    ELSIF ((x0 = TRUE) AND  (x1 = TRUE) AND  (x2 = FALSE) AND  (t0.Q = FALSE)) THEN 
        cstate58 := 2630; y0 := FALSE; y1 := FALSE; t0_start := FALSE; 
    ELSIF ((x0 = TRUE) AND  (x1 = TRUE) AND  (x2 = FALSE) AND  (t0.Q = TRUE)) THEN 
        cstate58 := 2626; y0 := FALSE; y1 := FALSE; t0_start := FALSE; 
    ELSIF ((x0 = TRUE) AND  (x1 = TRUE) AND  (x2 = TRUE) AND  (t0.Q = FALSE)) THEN 
        cstate58 := 2566; y0 := FALSE; y1 := FALSE; t0_start := TRUE; t0_up := FALSE; 
    ELSIF ((x0 = TRUE) AND  (x1 = TRUE) AND  (x2 = TRUE) AND  (t0.Q = TRUE)) THEN 
        cstate58 := 2562; y0 := FALSE; y1 := FALSE; t0_start := TRUE; t0_up := FALSE; 
    END_IF;
7428:
    IF ((x0 = FALSE) AND  (x1 = FALSE) AND  (x2 = FALSE) AND  (t0.Q = FALSE)) THEN 
        cstate58 := 7428; y0 := FALSE; y1 := FALSE; t0_start := FALSE; 
    ELSIF ((x0 = FALSE) AND  (x1 = FALSE) AND  (x2 = FALSE) AND  (t0.Q = TRUE)) THEN 
        cstate58 := 7370; y0 := FALSE; y1 := TRUE; t0_start := FALSE; 
    ELSIF ((x0 = FALSE) AND  (x1 = FALSE) AND  (x2 = TRUE) AND  (t0.Q = FALSE)) THEN 
        cstate58 := 7492; y0 := FALSE; y1 := FALSE; t0_start := TRUE; t0_up := FALSE; 
    ELSIF ((x0 = FALSE) AND  (x1 = FALSE) AND  (x2 = TRUE) AND  (t0.Q = TRUE)) THEN 
        cstate58 := 7500; y0 := FALSE; y1 := TRUE; t0_start := TRUE; t0_up := FALSE; 
    ELSIF ((x0 = FALSE) AND  (x1 = TRUE) AND  (x2 = FALSE) AND  (t0.Q = FALSE)) THEN 
        cstate58 := 6404; y0 := FALSE; y1 := FALSE; t0_start := FALSE; 
    ELSIF ((x0 = FALSE) AND  (x1 = TRUE) AND  (x2 = FALSE) AND  (t0.Q = TRUE)) THEN 
        cstate58 := 6338; y0 := FALSE; y1 := FALSE; t0_start := FALSE; 
    ELSIF ((x0 = FALSE) AND  (x1 = TRUE) AND  (x2 = TRUE) AND  (t0.Q = FALSE)) THEN 
        cstate58 := 6468; y0 := FALSE; y1 := FALSE; t0_start := TRUE; t0_up := FALSE; 
    ELSIF ((x0 = FALSE) AND  (x1 = TRUE) AND  (x2 = TRUE) AND  (t0.Q = TRUE)) THEN 
        cstate58 := 6466; y0 := FALSE; y1 := FALSE; t0_start := TRUE; t0_up := FALSE; 
    ELSIF ((x0 = TRUE) AND  (x1 = FALSE) AND  (x2 = FALSE) AND  (t0.Q = FALSE)) THEN 
        cstate58 := 5256; y0 := TRUE; y1 := FALSE; t0_start := FALSE; 
    ELSIF ((x0 = TRUE) AND  (x1 = FALSE) AND  (x2 = FALSE) AND  (t0.Q = TRUE)) THEN 
        cstate58 := 5186; y0 := TRUE; y1 := FALSE; t0_start := FALSE; 
    ELSIF ((x0 = TRUE) AND  (x1 = FALSE) AND  (x2 = TRUE) AND  (t0.Q = FALSE)) THEN 
        cstate58 := 3784; y0 := FALSE; y1 := FALSE; t0_start := TRUE; t0_up := FALSE; 
    ELSIF ((x0 = TRUE) AND  (x1 = FALSE) AND  (x2 = TRUE) AND  (t0.Q = TRUE)) THEN 
        cstate58 := 3778; y0 := FALSE; y1 := FALSE; t0_start := TRUE; t0_up := FALSE; 
    ELSIF ((x0 = TRUE) AND  (x1 = TRUE) AND  (x2 = FALSE) AND  (t0.Q = FALSE)) THEN 
        cstate58 := 4742; y0 := TRUE; y1 := FALSE; t0_start := FALSE; 
    ELSIF ((x0 = TRUE) AND  (x1 = TRUE) AND  (x2 = FALSE) AND  (t0.Q = TRUE)) THEN 
        cstate58 := 4674; y0 := TRUE; y1 := FALSE; t0_start := FALSE; 
    ELSIF ((x0 = TRUE) AND  (x1 = TRUE) AND  (x2 = TRUE) AND  (t0.Q = FALSE)) THEN 
        cstate58 := 2566; y0 := FALSE; y1 := FALSE; t0_start := TRUE; t0_up := FALSE; 
    ELSIF ((x0 = TRUE) AND  (x1 = TRUE) AND  (x2 = TRUE) AND  (t0.Q = TRUE)) THEN 
        cstate58 := 2562; y0 := FALSE; y1 := FALSE; t0_start := TRUE; t0_up := FALSE; 
    END_IF;
1304:
    IF ((x0 = FALSE) AND  (x1 = FALSE) AND  (x2 = FALSE) AND  (t0.Q = FALSE)) THEN 
        cstate58 := 1304; y0 := FALSE; y1 := TRUE; t0_start := FALSE; 
    ELSIF ((x0 = FALSE) AND  (x1 = FALSE) AND  (x2 = FALSE) AND  (t0.Q = TRUE)) THEN 
        cstate58 := 1226; y0 := FALSE; y1 := TRUE; t0_start := FALSE; 
    ELSIF ((x0 = FALSE) AND  (x1 = FALSE) AND  (x2 = TRUE) AND  (t0.Q = FALSE)) THEN 
        cstate58 := 1368; y0 := FALSE; y1 := TRUE; t0_start := TRUE; t0_up := FALSE; 
    ELSIF ((x0 = FALSE) AND  (x1 = FALSE) AND  (x2 = TRUE) AND  (t0.Q = TRUE)) THEN 
        cstate58 := 1356; y0 := FALSE; y1 := TRUE; t0_start := TRUE; t0_up := FALSE; 
    ELSIF ((x0 = FALSE) AND  (x1 = TRUE) AND  (x2 = FALSE) AND  (t0.Q = FALSE)) THEN 
        cstate58 := 1284; y0 := FALSE; y1 := FALSE; t0_start := FALSE; 
    ELSIF ((x0 = FALSE) AND  (x1 = TRUE) AND  (x2 = FALSE) AND  (t0.Q = TRUE)) THEN 
        cstate58 := 1218; y0 := FALSE; y1 := FALSE; t0_start := FALSE; 
    ELSIF ((x0 = FALSE) AND  (x1 = TRUE) AND  (x2 = TRUE) AND  (t0.Q = FALSE)) THEN 
        cstate58 := 1348; y0 := FALSE; y1 := FALSE; t0_start := TRUE; t0_up := FALSE; 
    ELSIF ((x0 = FALSE) AND  (x1 = TRUE) AND  (x2 = TRUE) AND  (t0.Q = TRUE)) THEN 
        cstate58 := 1346; y0 := FALSE; y1 := FALSE; t0_start := TRUE; t0_up := FALSE; 
    ELSIF ((x0 = TRUE) AND  (x1 = FALSE) AND  (x2 = FALSE) AND  (t0.Q = FALSE)) THEN 
        cstate58 := 5256; y0 := TRUE; y1 := FALSE; t0_start := FALSE; 
    ELSIF ((x0 = TRUE) AND  (x1 = FALSE) AND  (x2 = FALSE) AND  (t0.Q = TRUE)) THEN 
        cstate58 := 5186; y0 := TRUE; y1 := FALSE; t0_start := FALSE; 
    ELSIF ((x0 = TRUE) AND  (x1 = FALSE) AND  (x2 = TRUE) AND  (t0.Q = FALSE)) THEN 
        cstate58 := 3784; y0 := FALSE; y1 := FALSE; t0_start := TRUE; t0_up := FALSE; 
    ELSIF ((x0 = TRUE) AND  (x1 = FALSE) AND  (x2 = TRUE) AND  (t0.Q = TRUE)) THEN 
        cstate58 := 3778; y0 := FALSE; y1 := FALSE; t0_start := TRUE; t0_up := FALSE; 
    ELSIF ((x0 = TRUE) AND  (x1 = TRUE) AND  (x2 = FALSE) AND  (t0.Q = FALSE)) THEN 
        cstate58 := 4742; y0 := TRUE; y1 := FALSE; t0_start := FALSE; 
    ELSIF ((x0 = TRUE) AND  (x1 = TRUE) AND  (x2 = FALSE) AND  (t0.Q = TRUE)) THEN 
        cstate58 := 4674; y0 := TRUE; y1 := FALSE; t0_start := FALSE; 
    ELSIF ((x0 = TRUE) AND  (x1 = TRUE) AND  (x2 = TRUE) AND  (t0.Q = FALSE)) THEN 
        cstate58 := 2566; y0 := FALSE; y1 := FALSE; t0_start := TRUE; t0_up := FALSE; 
    ELSIF ((x0 = TRUE) AND  (x1 = TRUE) AND  (x2 = TRUE) AND  (t0.Q = TRUE)) THEN 
        cstate58 := 2562; y0 := FALSE; y1 := FALSE; t0_start := TRUE; t0_up := FALSE; 
    END_IF;
2824:
    IF ((x0 = FALSE) AND  (x1 = FALSE) AND  (x2 = FALSE) AND  (t0.Q = FALSE)) THEN 
        cstate58 := 6340; y0 := FALSE; y1 := FALSE; t0_start := FALSE; 
    ELSIF ((x0 = FALSE) AND  (x1 = FALSE) AND  (x2 = FALSE) AND  (t0.Q = TRUE)) THEN 
        cstate58 := 6354; y0 := FALSE; y1 := TRUE; t0_start := FALSE; 
    ELSIF ((x0 = FALSE) AND  (x1 = FALSE) AND  (x2 = TRUE) AND  (t0.Q = FALSE)) THEN 
        cstate58 := 6532; y0 := FALSE; y1 := FALSE; t0_start := FALSE; 
    ELSIF ((x0 = FALSE) AND  (x1 = FALSE) AND  (x2 = TRUE) AND  (t0.Q = TRUE)) THEN 
        cstate58 := 6546; y0 := FALSE; y1 := TRUE; t0_start := FALSE; 
    ELSIF ((x0 = FALSE) AND  (x1 = TRUE) AND  (x2 = FALSE) AND  (t0.Q = FALSE)) THEN 
        cstate58 := 6340; y0 := FALSE; y1 := FALSE; t0_start := FALSE; 
    ELSIF ((x0 = FALSE) AND  (x1 = TRUE) AND  (x2 = FALSE) AND  (t0.Q = TRUE)) THEN 
        cstate58 := 6338; y0 := FALSE; y1 := FALSE; t0_start := FALSE; 
    ELSIF ((x0 = FALSE) AND  (x1 = TRUE) AND  (x2 = TRUE) AND  (t0.Q = FALSE)) THEN 
        cstate58 := 6532; y0 := FALSE; y1 := FALSE; t0_start := FALSE; 
    ELSIF ((x0 = FALSE) AND  (x1 = TRUE) AND  (x2 = TRUE) AND  (t0.Q = TRUE)) THEN 
        cstate58 := 6530; y0 := FALSE; y1 := FALSE; t0_start := FALSE; 
    ELSIF ((x0 = TRUE) AND  (x1 = FALSE) AND  (x2 = FALSE) AND  (t0.Q = FALSE)) THEN 
        cstate58 := 2120; y0 := FALSE; y1 := FALSE; t0_start := FALSE; 
    ELSIF ((x0 = TRUE) AND  (x1 = FALSE) AND  (x2 = FALSE) AND  (t0.Q = TRUE)) THEN 
        cstate58 := 2114; y0 := FALSE; y1 := FALSE; t0_start := FALSE; 
    ELSIF ((x0 = TRUE) AND  (x1 = FALSE) AND  (x2 = TRUE) AND  (t0.Q = FALSE)) THEN 
        cstate58 := 2824; y0 := FALSE; y1 := FALSE; t0_start := FALSE; 
    ELSIF ((x0 = TRUE) AND  (x1 = FALSE) AND  (x2 = TRUE) AND  (t0.Q = TRUE)) THEN 
        cstate58 := 2818; y0 := FALSE; y1 := FALSE; t0_start := FALSE; 
    ELSIF ((x0 = TRUE) AND  (x1 = TRUE) AND  (x2 = FALSE) AND  (t0.Q = FALSE)) THEN 
        cstate58 := 2630; y0 := FALSE; y1 := FALSE; t0_start := FALSE; 
    ELSIF ((x0 = TRUE) AND  (x1 = TRUE) AND  (x2 = FALSE) AND  (t0.Q = TRUE)) THEN 
        cstate58 := 2626; y0 := FALSE; y1 := FALSE; t0_start := FALSE; 
    ELSIF ((x0 = TRUE) AND  (x1 = TRUE) AND  (x2 = TRUE) AND  (t0.Q = FALSE)) THEN 
        cstate58 := 2502; y0 := FALSE; y1 := FALSE; t0_start := FALSE; 
    ELSIF ((x0 = TRUE) AND  (x1 = TRUE) AND  (x2 = TRUE) AND  (t0.Q = TRUE)) THEN 
        cstate58 := 2498; y0 := FALSE; y1 := FALSE; t0_start := FALSE; 
    END_IF;
6480:
    IF ((x0 = FALSE) AND  (x1 = FALSE) AND  (x2 = FALSE) AND  (t0.Q = FALSE)) THEN 
        cstate58 := 6428; y0 := FALSE; y1 := TRUE; t0_start := FALSE; 
    ELSIF ((x0 = FALSE) AND  (x1 = FALSE) AND  (x2 = FALSE) AND  (t0.Q = TRUE)) THEN 
        cstate58 := 6350; y0 := FALSE; y1 := TRUE; t0_start := FALSE; 
    ELSIF ((x0 = FALSE) AND  (x1 = FALSE) AND  (x2 = TRUE) AND  (t0.Q = FALSE)) THEN 
        cstate58 := 6492; y0 := FALSE; y1 := TRUE; t0_start := FALSE; 
    ELSIF ((x0 = FALSE) AND  (x1 = FALSE) AND  (x2 = TRUE) AND  (t0.Q = TRUE)) THEN 
        cstate58 := 6542; y0 := FALSE; y1 := TRUE; t0_start := FALSE; 
    ELSIF ((x0 = FALSE) AND  (x1 = TRUE) AND  (x2 = FALSE) AND  (t0.Q = FALSE)) THEN 
        cstate58 := 6404; y0 := FALSE; y1 := FALSE; t0_start := FALSE; 
    ELSIF ((x0 = FALSE) AND  (x1 = TRUE) AND  (x2 = FALSE) AND  (t0.Q = TRUE)) THEN 
        cstate58 := 6338; y0 := FALSE; y1 := FALSE; t0_start := FALSE; 
    ELSIF ((x0 = FALSE) AND  (x1 = TRUE) AND  (x2 = TRUE) AND  (t0.Q = FALSE)) THEN 
        cstate58 := 6468; y0 := FALSE; y1 := FALSE; t0_start := FALSE; 
    ELSIF ((x0 = FALSE) AND  (x1 = TRUE) AND  (x2 = TRUE) AND  (t0.Q = TRUE)) THEN 
        cstate58 := 6530; y0 := FALSE; y1 := FALSE; t0_start := FALSE; 
    ELSIF ((x0 = TRUE) AND  (x1 = FALSE) AND  (x2 = FALSE) AND  (t0.Q = FALSE)) THEN 
        cstate58 := 4232; y0 := TRUE; y1 := FALSE; t0_start := FALSE; 
    ELSIF ((x0 = TRUE) AND  (x1 = FALSE) AND  (x2 = FALSE) AND  (t0.Q = TRUE)) THEN 
        cstate58 := 4162; y0 := TRUE; y1 := FALSE; t0_start := FALSE; 
    ELSIF ((x0 = TRUE) AND  (x1 = FALSE) AND  (x2 = TRUE) AND  (t0.Q = FALSE)) THEN 
        cstate58 := 2760; y0 := FALSE; y1 := FALSE; t0_start := FALSE; 
    ELSIF ((x0 = TRUE) AND  (x1 = FALSE) AND  (x2 = TRUE) AND  (t0.Q = TRUE)) THEN 
        cstate58 := 2818; y0 := FALSE; y1 := FALSE; t0_start := FALSE; 
    ELSIF ((x0 = TRUE) AND  (x1 = TRUE) AND  (x2 = FALSE) AND  (t0.Q = FALSE)) THEN 
        cstate58 := 4742; y0 := TRUE; y1 := FALSE; t0_start := FALSE; 
    ELSIF ((x0 = TRUE) AND  (x1 = TRUE) AND  (x2 = FALSE) AND  (t0.Q = TRUE)) THEN 
        cstate58 := 4674; y0 := TRUE; y1 := FALSE; t0_start := FALSE; 
    ELSIF ((x0 = TRUE) AND  (x1 = TRUE) AND  (x2 = TRUE) AND  (t0.Q = FALSE)) THEN 
        cstate58 := 2566; y0 := FALSE; y1 := FALSE; t0_start := FALSE; 
    ELSIF ((x0 = TRUE) AND  (x1 = TRUE) AND  (x2 = TRUE) AND  (t0.Q = TRUE)) THEN 
        cstate58 := 2498; y0 := FALSE; y1 := FALSE; t0_start := FALSE; 
    END_IF;
6484:
    IF ((x0 = FALSE) AND  (x1 = FALSE) AND  (x2 = FALSE) AND  (t0.Q = FALSE)) THEN 
        cstate58 := 6432; y0 := FALSE; y1 := TRUE; t0_start := FALSE; 
    ELSIF ((x0 = FALSE) AND  (x1 = FALSE) AND  (x2 = FALSE) AND  (t0.Q = TRUE)) THEN 
        cstate58 := 6354; y0 := FALSE; y1 := TRUE; t0_start := FALSE; 
    ELSIF ((x0 = FALSE) AND  (x1 = FALSE) AND  (x2 = TRUE) AND  (t0.Q = FALSE)) THEN 
        cstate58 := 6496; y0 := FALSE; y1 := TRUE; t0_start := FALSE; 
    ELSIF ((x0 = FALSE) AND  (x1 = FALSE) AND  (x2 = TRUE) AND  (t0.Q = TRUE)) THEN 
        cstate58 := 6546; y0 := FALSE; y1 := TRUE; t0_start := FALSE; 
    ELSIF ((x0 = FALSE) AND  (x1 = TRUE) AND  (x2 = FALSE) AND  (t0.Q = FALSE)) THEN 
        cstate58 := 6404; y0 := FALSE; y1 := FALSE; t0_start := FALSE; 
    ELSIF ((x0 = FALSE) AND  (x1 = TRUE) AND  (x2 = FALSE) AND  (t0.Q = TRUE)) THEN 
        cstate58 := 6338; y0 := FALSE; y1 := FALSE; t0_start := FALSE; 
    ELSIF ((x0 = FALSE) AND  (x1 = TRUE) AND  (x2 = TRUE) AND  (t0.Q = FALSE)) THEN 
        cstate58 := 6468; y0 := FALSE; y1 := FALSE; t0_start := FALSE; 
    ELSIF ((x0 = FALSE) AND  (x1 = TRUE) AND  (x2 = TRUE) AND  (t0.Q = TRUE)) THEN 
        cstate58 := 6530; y0 := FALSE; y1 := FALSE; t0_start := FALSE; 
    ELSIF ((x0 = TRUE) AND  (x1 = FALSE) AND  (x2 = FALSE) AND  (t0.Q = FALSE)) THEN 
        cstate58 := 4232; y0 := TRUE; y1 := FALSE; t0_start := FALSE; 
    ELSIF ((x0 = TRUE) AND  (x1 = FALSE) AND  (x2 = FALSE) AND  (t0.Q = TRUE)) THEN 
        cstate58 := 4162; y0 := TRUE; y1 := FALSE; t0_start := FALSE; 
    ELSIF ((x0 = TRUE) AND  (x1 = FALSE) AND  (x2 = TRUE) AND  (t0.Q = FALSE)) THEN 
        cstate58 := 2760; y0 := FALSE; y1 := FALSE; t0_start := FALSE; 
    ELSIF ((x0 = TRUE) AND  (x1 = FALSE) AND  (x2 = TRUE) AND  (t0.Q = TRUE)) THEN 
        cstate58 := 2818; y0 := FALSE; y1 := FALSE; t0_start := FALSE; 
    ELSIF ((x0 = TRUE) AND  (x1 = TRUE) AND  (x2 = FALSE) AND  (t0.Q = FALSE)) THEN 
        cstate58 := 4742; y0 := TRUE; y1 := FALSE; t0_start := FALSE; 
    ELSIF ((x0 = TRUE) AND  (x1 = TRUE) AND  (x2 = FALSE) AND  (t0.Q = TRUE)) THEN 
        cstate58 := 4674; y0 := TRUE; y1 := FALSE; t0_start := FALSE; 
    ELSIF ((x0 = TRUE) AND  (x1 = TRUE) AND  (x2 = TRUE) AND  (t0.Q = FALSE)) THEN 
        cstate58 := 2566; y0 := FALSE; y1 := FALSE; t0_start := FALSE; 
    ELSIF ((x0 = TRUE) AND  (x1 = TRUE) AND  (x2 = TRUE) AND  (t0.Q = TRUE)) THEN 
        cstate58 := 2498; y0 := FALSE; y1 := FALSE; t0_start := FALSE; 
    END_IF;
2184:
    IF ((x0 = FALSE) AND  (x1 = FALSE) AND  (x2 = FALSE) AND  (t0.Q = FALSE)) THEN 
        cstate58 := 6404; y0 := FALSE; y1 := FALSE; t0_start := FALSE; 
    ELSIF ((x0 = FALSE) AND  (x1 = FALSE) AND  (x2 = FALSE) AND  (t0.Q = TRUE)) THEN 
        cstate58 := 6354; y0 := FALSE; y1 := TRUE; t0_start := FALSE; 
    ELSIF ((x0 = FALSE) AND  (x1 = FALSE) AND  (x2 = TRUE) AND  (t0.Q = FALSE)) THEN 
        cstate58 := 6468; y0 := FALSE; y1 := FALSE; t0_start := TRUE; t0_up := FALSE; 
    ELSIF ((x0 = FALSE) AND  (x1 = FALSE) AND  (x2 = TRUE) AND  (t0.Q = TRUE)) THEN 
        cstate58 := 6484; y0 := FALSE; y1 := TRUE; t0_start := TRUE; t0_up := FALSE; 
    ELSIF ((x0 = FALSE) AND  (x1 = TRUE) AND  (x2 = FALSE) AND  (t0.Q = FALSE)) THEN 
        cstate58 := 6404; y0 := FALSE; y1 := FALSE; t0_start := FALSE; 
    ELSIF ((x0 = FALSE) AND  (x1 = TRUE) AND  (x2 = FALSE) AND  (t0.Q = TRUE)) THEN 
        cstate58 := 6338; y0 := FALSE; y1 := FALSE; t0_start := FALSE; 
    ELSIF ((x0 = FALSE) AND  (x1 = TRUE) AND  (x2 = TRUE) AND  (t0.Q = FALSE)) THEN 
        cstate58 := 6468; y0 := FALSE; y1 := FALSE; t0_start := TRUE; t0_up := FALSE; 
    ELSIF ((x0 = FALSE) AND  (x1 = TRUE) AND  (x2 = TRUE) AND  (t0.Q = TRUE)) THEN 
        cstate58 := 6466; y0 := FALSE; y1 := FALSE; t0_start := TRUE; t0_up := FALSE; 
    ELSIF ((x0 = TRUE) AND  (x1 = FALSE) AND  (x2 = FALSE) AND  (t0.Q = FALSE)) THEN 
        cstate58 := 2184; y0 := FALSE; y1 := FALSE; t0_start := FALSE; 
    ELSIF ((x0 = TRUE) AND  (x1 = FALSE) AND  (x2 = FALSE) AND  (t0.Q = TRUE)) THEN 
        cstate58 := 2114; y0 := FALSE; y1 := FALSE; t0_start := FALSE; 
    ELSIF ((x0 = TRUE) AND  (x1 = FALSE) AND  (x2 = TRUE) AND  (t0.Q = FALSE)) THEN 
        cstate58 := 2760; y0 := FALSE; y1 := FALSE; t0_start := TRUE; t0_up := FALSE; 
    ELSIF ((x0 = TRUE) AND  (x1 = FALSE) AND  (x2 = TRUE) AND  (t0.Q = TRUE)) THEN 
        cstate58 := 2754; y0 := FALSE; y1 := FALSE; t0_start := TRUE; t0_up := FALSE; 
    ELSIF ((x0 = TRUE) AND  (x1 = TRUE) AND  (x2 = FALSE) AND  (t0.Q = FALSE)) THEN 
        cstate58 := 2694; y0 := FALSE; y1 := FALSE; t0_start := FALSE; 
    ELSIF ((x0 = TRUE) AND  (x1 = TRUE) AND  (x2 = FALSE) AND  (t0.Q = TRUE)) THEN 
        cstate58 := 2626; y0 := FALSE; y1 := FALSE; t0_start := FALSE; 
    ELSIF ((x0 = TRUE) AND  (x1 = TRUE) AND  (x2 = TRUE) AND  (t0.Q = FALSE)) THEN 
        cstate58 := 2566; y0 := FALSE; y1 := FALSE; t0_start := TRUE; t0_up := FALSE; 
    ELSIF ((x0 = TRUE) AND  (x1 = TRUE) AND  (x2 = TRUE) AND  (t0.Q = TRUE)) THEN 
        cstate58 := 2562; y0 := FALSE; y1 := FALSE; t0_start := TRUE; t0_up := FALSE; 
    END_IF;
6488:
    IF ((x0 = FALSE) AND  (x1 = FALSE) AND  (x2 = FALSE) AND  (t0.Q = FALSE)) THEN 
        cstate58 := 6424; y0 := FALSE; y1 := TRUE; t0_start := FALSE; 
    ELSIF ((x0 = FALSE) AND  (x1 = FALSE) AND  (x2 = FALSE) AND  (t0.Q = TRUE)) THEN 
        cstate58 := 6346; y0 := FALSE; y1 := TRUE; t0_start := FALSE; 
    ELSIF ((x0 = FALSE) AND  (x1 = FALSE) AND  (x2 = TRUE) AND  (t0.Q = FALSE)) THEN 
        cstate58 := 6488; y0 := FALSE; y1 := TRUE; t0_start := FALSE; 
    ELSIF ((x0 = FALSE) AND  (x1 = FALSE) AND  (x2 = TRUE) AND  (t0.Q = TRUE)) THEN 
        cstate58 := 6538; y0 := FALSE; y1 := TRUE; t0_start := FALSE; 
    ELSIF ((x0 = FALSE) AND  (x1 = TRUE) AND  (x2 = FALSE) AND  (t0.Q = FALSE)) THEN 
        cstate58 := 6404; y0 := FALSE; y1 := FALSE; t0_start := FALSE; 
    ELSIF ((x0 = FALSE) AND  (x1 = TRUE) AND  (x2 = FALSE) AND  (t0.Q = TRUE)) THEN 
        cstate58 := 6338; y0 := FALSE; y1 := FALSE; t0_start := FALSE; 
    ELSIF ((x0 = FALSE) AND  (x1 = TRUE) AND  (x2 = TRUE) AND  (t0.Q = FALSE)) THEN 
        cstate58 := 6468; y0 := FALSE; y1 := FALSE; t0_start := FALSE; 
    ELSIF ((x0 = FALSE) AND  (x1 = TRUE) AND  (x2 = TRUE) AND  (t0.Q = TRUE)) THEN 
        cstate58 := 6530; y0 := FALSE; y1 := FALSE; t0_start := FALSE; 
    ELSIF ((x0 = TRUE) AND  (x1 = FALSE) AND  (x2 = FALSE) AND  (t0.Q = FALSE)) THEN 
        cstate58 := 4232; y0 := TRUE; y1 := FALSE; t0_start := FALSE; 
    ELSIF ((x0 = TRUE) AND  (x1 = FALSE) AND  (x2 = FALSE) AND  (t0.Q = TRUE)) THEN 
        cstate58 := 4162; y0 := TRUE; y1 := FALSE; t0_start := FALSE; 
    ELSIF ((x0 = TRUE) AND  (x1 = FALSE) AND  (x2 = TRUE) AND  (t0.Q = FALSE)) THEN 
        cstate58 := 2760; y0 := FALSE; y1 := FALSE; t0_start := FALSE; 
    ELSIF ((x0 = TRUE) AND  (x1 = FALSE) AND  (x2 = TRUE) AND  (t0.Q = TRUE)) THEN 
        cstate58 := 2818; y0 := FALSE; y1 := FALSE; t0_start := FALSE; 
    ELSIF ((x0 = TRUE) AND  (x1 = TRUE) AND  (x2 = FALSE) AND  (t0.Q = FALSE)) THEN 
        cstate58 := 4742; y0 := TRUE; y1 := FALSE; t0_start := FALSE; 
    ELSIF ((x0 = TRUE) AND  (x1 = TRUE) AND  (x2 = FALSE) AND  (t0.Q = TRUE)) THEN 
        cstate58 := 4674; y0 := TRUE; y1 := FALSE; t0_start := FALSE; 
    ELSIF ((x0 = TRUE) AND  (x1 = TRUE) AND  (x2 = TRUE) AND  (t0.Q = FALSE)) THEN 
        cstate58 := 2566; y0 := FALSE; y1 := FALSE; t0_start := FALSE; 
    ELSIF ((x0 = TRUE) AND  (x1 = TRUE) AND  (x2 = TRUE) AND  (t0.Q = TRUE)) THEN 
        cstate58 := 2498; y0 := FALSE; y1 := FALSE; t0_start := FALSE; 
    END_IF;
6466:
    IF ((x0 = FALSE) AND  (x1 = FALSE) AND  (x2 = FALSE) AND  (t0.Q = FALSE)) THEN 
        cstate58 := 6404; y0 := FALSE; y1 := FALSE; t0_start := FALSE; 
    ELSIF ((x0 = FALSE) AND  (x1 = FALSE) AND  (x2 = FALSE) AND  (t0.Q = TRUE)) THEN 
        cstate58 := 6338; y0 := FALSE; y1 := FALSE; t0_start := FALSE; 
    ELSIF ((x0 = FALSE) AND  (x1 = FALSE) AND  (x2 = TRUE) AND  (t0.Q = FALSE)) THEN 
        cstate58 := 6468; y0 := FALSE; y1 := FALSE; t0_start := FALSE; 
    ELSIF ((x0 = FALSE) AND  (x1 = FALSE) AND  (x2 = TRUE) AND  (t0.Q = TRUE)) THEN 
        cstate58 := 6530; y0 := FALSE; y1 := FALSE; t0_start := FALSE; 
    ELSIF ((x0 = FALSE) AND  (x1 = TRUE) AND  (x2 = FALSE) AND  (t0.Q = FALSE)) THEN 
        cstate58 := 6404; y0 := FALSE; y1 := FALSE; t0_start := FALSE; 
    ELSIF ((x0 = FALSE) AND  (x1 = TRUE) AND  (x2 = FALSE) AND  (t0.Q = TRUE)) THEN 
        cstate58 := 6338; y0 := FALSE; y1 := FALSE; t0_start := FALSE; 
    ELSIF ((x0 = FALSE) AND  (x1 = TRUE) AND  (x2 = TRUE) AND  (t0.Q = FALSE)) THEN 
        cstate58 := 6468; y0 := FALSE; y1 := FALSE; t0_start := FALSE; 
    ELSIF ((x0 = FALSE) AND  (x1 = TRUE) AND  (x2 = TRUE) AND  (t0.Q = TRUE)) THEN 
        cstate58 := 6530; y0 := FALSE; y1 := FALSE; t0_start := FALSE; 
    ELSIF ((x0 = TRUE) AND  (x1 = FALSE) AND  (x2 = FALSE) AND  (t0.Q = FALSE)) THEN 
        cstate58 := 4232; y0 := TRUE; y1 := FALSE; t0_start := FALSE; 
    ELSIF ((x0 = TRUE) AND  (x1 = FALSE) AND  (x2 = FALSE) AND  (t0.Q = TRUE)) THEN 
        cstate58 := 4162; y0 := TRUE; y1 := FALSE; t0_start := FALSE; 
    ELSIF ((x0 = TRUE) AND  (x1 = FALSE) AND  (x2 = TRUE) AND  (t0.Q = FALSE)) THEN 
        cstate58 := 2760; y0 := FALSE; y1 := FALSE; t0_start := FALSE; 
    ELSIF ((x0 = TRUE) AND  (x1 = FALSE) AND  (x2 = TRUE) AND  (t0.Q = TRUE)) THEN 
        cstate58 := 2818; y0 := FALSE; y1 := FALSE; t0_start := FALSE; 
    ELSIF ((x0 = TRUE) AND  (x1 = TRUE) AND  (x2 = FALSE) AND  (t0.Q = FALSE)) THEN 
        cstate58 := 4742; y0 := TRUE; y1 := FALSE; t0_start := FALSE; 
    ELSIF ((x0 = TRUE) AND  (x1 = TRUE) AND  (x2 = FALSE) AND  (t0.Q = TRUE)) THEN 
        cstate58 := 4674; y0 := TRUE; y1 := FALSE; t0_start := FALSE; 
    ELSIF ((x0 = TRUE) AND  (x1 = TRUE) AND  (x2 = TRUE) AND  (t0.Q = FALSE)) THEN 
        cstate58 := 2566; y0 := FALSE; y1 := FALSE; t0_start := FALSE; 
    ELSIF ((x0 = TRUE) AND  (x1 = TRUE) AND  (x2 = TRUE) AND  (t0.Q = TRUE)) THEN 
        cstate58 := 2498; y0 := FALSE; y1 := FALSE; t0_start := FALSE; 
    END_IF;
9410:
    IF ((x0 = FALSE) AND  (x1 = FALSE) AND  (x2 = FALSE) AND  (t0.Q = FALSE)) THEN 
        cstate58 := 9412; y0 := TRUE; y1 := FALSE; t0_start := FALSE; 
    ELSIF ((x0 = FALSE) AND  (x1 = FALSE) AND  (x2 = FALSE) AND  (t0.Q = TRUE)) THEN 
        cstate58 := 9410; y0 := TRUE; y1 := FALSE; t0_start := FALSE; 
    ELSIF ((x0 = FALSE) AND  (x1 = FALSE) AND  (x2 = TRUE) AND  (t0.Q = FALSE)) THEN 
        cstate58 := 7492; y0 := FALSE; y1 := FALSE; t0_start := TRUE; t0_up := FALSE; 
    ELSIF ((x0 = FALSE) AND  (x1 = FALSE) AND  (x2 = TRUE) AND  (t0.Q = TRUE)) THEN 
        cstate58 := 7490; y0 := FALSE; y1 := FALSE; t0_start := TRUE; t0_up := FALSE; 
    ELSIF ((x0 = FALSE) AND  (x1 = TRUE) AND  (x2 = FALSE) AND  (t0.Q = FALSE)) THEN 
        cstate58 := 8388; y0 := TRUE; y1 := FALSE; t0_start := FALSE; 
    ELSIF ((x0 = FALSE) AND  (x1 = TRUE) AND  (x2 = FALSE) AND  (t0.Q = TRUE)) THEN 
        cstate58 := 8386; y0 := TRUE; y1 := FALSE; t0_start := FALSE; 
    ELSIF ((x0 = FALSE) AND  (x1 = TRUE) AND  (x2 = TRUE) AND  (t0.Q = FALSE)) THEN 
        cstate58 := 6468; y0 := FALSE; y1 := FALSE; t0_start := TRUE; t0_up := FALSE; 
    ELSIF ((x0 = FALSE) AND  (x1 = TRUE) AND  (x2 = TRUE) AND  (t0.Q = TRUE)) THEN 
        cstate58 := 6466; y0 := FALSE; y1 := FALSE; t0_start := TRUE; t0_up := FALSE; 
    ELSIF ((x0 = TRUE) AND  (x1 = FALSE) AND  (x2 = FALSE) AND  (t0.Q = FALSE)) THEN 
        cstate58 := 5192; y0 := TRUE; y1 := FALSE; t0_start := FALSE; 
    ELSIF ((x0 = TRUE) AND  (x1 = FALSE) AND  (x2 = FALSE) AND  (t0.Q = TRUE)) THEN 
        cstate58 := 5186; y0 := TRUE; y1 := FALSE; t0_start := FALSE; 
    ELSIF ((x0 = TRUE) AND  (x1 = FALSE) AND  (x2 = TRUE) AND  (t0.Q = FALSE)) THEN 
        cstate58 := 3784; y0 := FALSE; y1 := FALSE; t0_start := TRUE; t0_up := FALSE; 
    ELSIF ((x0 = TRUE) AND  (x1 = FALSE) AND  (x2 = TRUE) AND  (t0.Q = TRUE)) THEN 
        cstate58 := 3778; y0 := FALSE; y1 := FALSE; t0_start := TRUE; t0_up := FALSE; 
    ELSIF ((x0 = TRUE) AND  (x1 = TRUE) AND  (x2 = FALSE) AND  (t0.Q = FALSE)) THEN 
        cstate58 := 4678; y0 := TRUE; y1 := FALSE; t0_start := FALSE; 
    ELSIF ((x0 = TRUE) AND  (x1 = TRUE) AND  (x2 = FALSE) AND  (t0.Q = TRUE)) THEN 
        cstate58 := 4674; y0 := TRUE; y1 := FALSE; t0_start := FALSE; 
    ELSIF ((x0 = TRUE) AND  (x1 = TRUE) AND  (x2 = TRUE) AND  (t0.Q = FALSE)) THEN 
        cstate58 := 2566; y0 := FALSE; y1 := FALSE; t0_start := TRUE; t0_up := FALSE; 
    ELSIF ((x0 = TRUE) AND  (x1 = TRUE) AND  (x2 = TRUE) AND  (t0.Q = TRUE)) THEN 
        cstate58 := 2562; y0 := FALSE; y1 := FALSE; t0_start := TRUE; t0_up := FALSE; 
    END_IF;
2818:
    IF ((x0 = FALSE) AND  (x1 = FALSE) AND  (x2 = FALSE) AND  (t0.Q = FALSE)) THEN 
        cstate58 := 6340; y0 := FALSE; y1 := FALSE; t0_start := FALSE; 
    ELSIF ((x0 = FALSE) AND  (x1 = FALSE) AND  (x2 = FALSE) AND  (t0.Q = TRUE)) THEN 
        cstate58 := 6338; y0 := FALSE; y1 := FALSE; t0_start := FALSE; 
    ELSIF ((x0 = FALSE) AND  (x1 = FALSE) AND  (x2 = TRUE) AND  (t0.Q = FALSE)) THEN 
        cstate58 := 6532; y0 := FALSE; y1 := FALSE; t0_start := FALSE; 
    ELSIF ((x0 = FALSE) AND  (x1 = FALSE) AND  (x2 = TRUE) AND  (t0.Q = TRUE)) THEN 
        cstate58 := 6530; y0 := FALSE; y1 := FALSE; t0_start := FALSE; 
    ELSIF ((x0 = FALSE) AND  (x1 = TRUE) AND  (x2 = FALSE) AND  (t0.Q = FALSE)) THEN 
        cstate58 := 6340; y0 := FALSE; y1 := FALSE; t0_start := FALSE; 
    ELSIF ((x0 = FALSE) AND  (x1 = TRUE) AND  (x2 = FALSE) AND  (t0.Q = TRUE)) THEN 
        cstate58 := 6338; y0 := FALSE; y1 := FALSE; t0_start := FALSE; 
    ELSIF ((x0 = FALSE) AND  (x1 = TRUE) AND  (x2 = TRUE) AND  (t0.Q = FALSE)) THEN 
        cstate58 := 6532; y0 := FALSE; y1 := FALSE; t0_start := FALSE; 
    ELSIF ((x0 = FALSE) AND  (x1 = TRUE) AND  (x2 = TRUE) AND  (t0.Q = TRUE)) THEN 
        cstate58 := 6530; y0 := FALSE; y1 := FALSE; t0_start := FALSE; 
    ELSIF ((x0 = TRUE) AND  (x1 = FALSE) AND  (x2 = FALSE) AND  (t0.Q = FALSE)) THEN 
        cstate58 := 2120; y0 := FALSE; y1 := FALSE; t0_start := FALSE; 
    ELSIF ((x0 = TRUE) AND  (x1 = FALSE) AND  (x2 = FALSE) AND  (t0.Q = TRUE)) THEN 
        cstate58 := 2114; y0 := FALSE; y1 := FALSE; t0_start := FALSE; 
    ELSIF ((x0 = TRUE) AND  (x1 = FALSE) AND  (x2 = TRUE) AND  (t0.Q = FALSE)) THEN 
        cstate58 := 2824; y0 := FALSE; y1 := FALSE; t0_start := FALSE; 
    ELSIF ((x0 = TRUE) AND  (x1 = FALSE) AND  (x2 = TRUE) AND  (t0.Q = TRUE)) THEN 
        cstate58 := 2818; y0 := FALSE; y1 := FALSE; t0_start := FALSE; 
    ELSIF ((x0 = TRUE) AND  (x1 = TRUE) AND  (x2 = FALSE) AND  (t0.Q = FALSE)) THEN 
        cstate58 := 2630; y0 := FALSE; y1 := FALSE; t0_start := FALSE; 
    ELSIF ((x0 = TRUE) AND  (x1 = TRUE) AND  (x2 = FALSE) AND  (t0.Q = TRUE)) THEN 
        cstate58 := 2626; y0 := FALSE; y1 := FALSE; t0_start := FALSE; 
    ELSIF ((x0 = TRUE) AND  (x1 = TRUE) AND  (x2 = TRUE) AND  (t0.Q = FALSE)) THEN 
        cstate58 := 2502; y0 := FALSE; y1 := FALSE; t0_start := FALSE; 
    ELSIF ((x0 = TRUE) AND  (x1 = TRUE) AND  (x2 = TRUE) AND  (t0.Q = TRUE)) THEN 
        cstate58 := 2498; y0 := FALSE; y1 := FALSE; t0_start := FALSE; 
    END_IF;
9412:
    IF ((x0 = FALSE) AND  (x1 = FALSE) AND  (x2 = FALSE) AND  (t0.Q = FALSE)) THEN 
        cstate58 := 9412; y0 := TRUE; y1 := FALSE; t0_start := FALSE; 
    ELSIF ((x0 = FALSE) AND  (x1 = FALSE) AND  (x2 = FALSE) AND  (t0.Q = TRUE)) THEN 
        cstate58 := 9410; y0 := TRUE; y1 := FALSE; t0_start := FALSE; 
    ELSIF ((x0 = FALSE) AND  (x1 = FALSE) AND  (x2 = TRUE) AND  (t0.Q = FALSE)) THEN 
        cstate58 := 7492; y0 := FALSE; y1 := FALSE; t0_start := TRUE; t0_up := FALSE; 
    ELSIF ((x0 = FALSE) AND  (x1 = FALSE) AND  (x2 = TRUE) AND  (t0.Q = TRUE)) THEN 
        cstate58 := 7500; y0 := FALSE; y1 := TRUE; t0_start := TRUE; t0_up := FALSE; 
    ELSIF ((x0 = FALSE) AND  (x1 = TRUE) AND  (x2 = FALSE) AND  (t0.Q = FALSE)) THEN 
        cstate58 := 8388; y0 := TRUE; y1 := FALSE; t0_start := FALSE; 
    ELSIF ((x0 = FALSE) AND  (x1 = TRUE) AND  (x2 = FALSE) AND  (t0.Q = TRUE)) THEN 
        cstate58 := 8386; y0 := TRUE; y1 := FALSE; t0_start := FALSE; 
    ELSIF ((x0 = FALSE) AND  (x1 = TRUE) AND  (x2 = TRUE) AND  (t0.Q = FALSE)) THEN 
        cstate58 := 6468; y0 := FALSE; y1 := FALSE; t0_start := TRUE; t0_up := FALSE; 
    ELSIF ((x0 = FALSE) AND  (x1 = TRUE) AND  (x2 = TRUE) AND  (t0.Q = TRUE)) THEN 
        cstate58 := 6466; y0 := FALSE; y1 := FALSE; t0_start := TRUE; t0_up := FALSE; 
    ELSIF ((x0 = TRUE) AND  (x1 = FALSE) AND  (x2 = FALSE) AND  (t0.Q = FALSE)) THEN 
        cstate58 := 5192; y0 := TRUE; y1 := FALSE; t0_start := FALSE; 
    ELSIF ((x0 = TRUE) AND  (x1 = FALSE) AND  (x2 = FALSE) AND  (t0.Q = TRUE)) THEN 
        cstate58 := 5186; y0 := TRUE; y1 := FALSE; t0_start := FALSE; 
    ELSIF ((x0 = TRUE) AND  (x1 = FALSE) AND  (x2 = TRUE) AND  (t0.Q = FALSE)) THEN 
        cstate58 := 3784; y0 := FALSE; y1 := FALSE; t0_start := TRUE; t0_up := FALSE; 
    ELSIF ((x0 = TRUE) AND  (x1 = FALSE) AND  (x2 = TRUE) AND  (t0.Q = TRUE)) THEN 
        cstate58 := 3778; y0 := FALSE; y1 := FALSE; t0_start := TRUE; t0_up := FALSE; 
    ELSIF ((x0 = TRUE) AND  (x1 = TRUE) AND  (x2 = FALSE) AND  (t0.Q = FALSE)) THEN 
        cstate58 := 4678; y0 := TRUE; y1 := FALSE; t0_start := FALSE; 
    ELSIF ((x0 = TRUE) AND  (x1 = TRUE) AND  (x2 = FALSE) AND  (t0.Q = TRUE)) THEN 
        cstate58 := 4674; y0 := TRUE; y1 := FALSE; t0_start := FALSE; 
    ELSIF ((x0 = TRUE) AND  (x1 = TRUE) AND  (x2 = TRUE) AND  (t0.Q = FALSE)) THEN 
        cstate58 := 2566; y0 := FALSE; y1 := FALSE; t0_start := TRUE; t0_up := FALSE; 
    ELSIF ((x0 = TRUE) AND  (x1 = TRUE) AND  (x2 = TRUE) AND  (t0.Q = TRUE)) THEN 
        cstate58 := 2562; y0 := FALSE; y1 := FALSE; t0_start := TRUE; t0_up := FALSE; 
    END_IF;
7456:
    IF ((x0 = FALSE) AND  (x1 = FALSE) AND  (x2 = FALSE) AND  (t0.Q = FALSE)) THEN 
        cstate58 := 7456; y0 := FALSE; y1 := TRUE; t0_start := FALSE; 
    ELSIF ((x0 = FALSE) AND  (x1 = FALSE) AND  (x2 = FALSE) AND  (t0.Q = TRUE)) THEN 
        cstate58 := 7378; y0 := FALSE; y1 := TRUE; t0_start := FALSE; 
    ELSIF ((x0 = FALSE) AND  (x1 = FALSE) AND  (x2 = TRUE) AND  (t0.Q = FALSE)) THEN 
        cstate58 := 7520; y0 := FALSE; y1 := TRUE; t0_start := TRUE; t0_up := FALSE; 
    ELSIF ((x0 = FALSE) AND  (x1 = FALSE) AND  (x2 = TRUE) AND  (t0.Q = TRUE)) THEN 
        cstate58 := 7508; y0 := FALSE; y1 := TRUE; t0_start := TRUE; t0_up := FALSE; 
    ELSIF ((x0 = FALSE) AND  (x1 = TRUE) AND  (x2 = FALSE) AND  (t0.Q = FALSE)) THEN 
        cstate58 := 6404; y0 := FALSE; y1 := FALSE; t0_start := FALSE; 
    ELSIF ((x0 = FALSE) AND  (x1 = TRUE) AND  (x2 = FALSE) AND  (t0.Q = TRUE)) THEN 
        cstate58 := 6338; y0 := FALSE; y1 := FALSE; t0_start := FALSE; 
    ELSIF ((x0 = FALSE) AND  (x1 = TRUE) AND  (x2 = TRUE) AND  (t0.Q = FALSE)) THEN 
        cstate58 := 6468; y0 := FALSE; y1 := FALSE; t0_start := TRUE; t0_up := FALSE; 
    ELSIF ((x0 = FALSE) AND  (x1 = TRUE) AND  (x2 = TRUE) AND  (t0.Q = TRUE)) THEN 
        cstate58 := 6466; y0 := FALSE; y1 := FALSE; t0_start := TRUE; t0_up := FALSE; 
    ELSIF ((x0 = TRUE) AND  (x1 = FALSE) AND  (x2 = FALSE) AND  (t0.Q = FALSE)) THEN 
        cstate58 := 5256; y0 := TRUE; y1 := FALSE; t0_start := FALSE; 
    ELSIF ((x0 = TRUE) AND  (x1 = FALSE) AND  (x2 = FALSE) AND  (t0.Q = TRUE)) THEN 
        cstate58 := 5186; y0 := TRUE; y1 := FALSE; t0_start := FALSE; 
    ELSIF ((x0 = TRUE) AND  (x1 = FALSE) AND  (x2 = TRUE) AND  (t0.Q = FALSE)) THEN 
        cstate58 := 3784; y0 := FALSE; y1 := FALSE; t0_start := TRUE; t0_up := FALSE; 
    ELSIF ((x0 = TRUE) AND  (x1 = FALSE) AND  (x2 = TRUE) AND  (t0.Q = TRUE)) THEN 
        cstate58 := 3778; y0 := FALSE; y1 := FALSE; t0_start := TRUE; t0_up := FALSE; 
    ELSIF ((x0 = TRUE) AND  (x1 = TRUE) AND  (x2 = FALSE) AND  (t0.Q = FALSE)) THEN 
        cstate58 := 4742; y0 := TRUE; y1 := FALSE; t0_start := FALSE; 
    ELSIF ((x0 = TRUE) AND  (x1 = TRUE) AND  (x2 = FALSE) AND  (t0.Q = TRUE)) THEN 
        cstate58 := 4674; y0 := TRUE; y1 := FALSE; t0_start := FALSE; 
    ELSIF ((x0 = TRUE) AND  (x1 = TRUE) AND  (x2 = TRUE) AND  (t0.Q = FALSE)) THEN 
        cstate58 := 2566; y0 := FALSE; y1 := FALSE; t0_start := TRUE; t0_up := FALSE; 
    ELSIF ((x0 = TRUE) AND  (x1 = TRUE) AND  (x2 = TRUE) AND  (t0.Q = TRUE)) THEN 
        cstate58 := 2562; y0 := FALSE; y1 := FALSE; t0_start := TRUE; t0_up := FALSE; 
    END_IF;
7448:
    IF ((x0 = FALSE) AND  (x1 = FALSE) AND  (x2 = FALSE) AND  (t0.Q = FALSE)) THEN 
        cstate58 := 7448; y0 := FALSE; y1 := TRUE; t0_start := FALSE; 
    ELSIF ((x0 = FALSE) AND  (x1 = FALSE) AND  (x2 = FALSE) AND  (t0.Q = TRUE)) THEN 
        cstate58 := 7370; y0 := FALSE; y1 := TRUE; t0_start := FALSE; 
    ELSIF ((x0 = FALSE) AND  (x1 = FALSE) AND  (x2 = TRUE) AND  (t0.Q = FALSE)) THEN 
        cstate58 := 7512; y0 := FALSE; y1 := TRUE; t0_start := TRUE; t0_up := FALSE; 
    ELSIF ((x0 = FALSE) AND  (x1 = FALSE) AND  (x2 = TRUE) AND  (t0.Q = TRUE)) THEN 
        cstate58 := 7500; y0 := FALSE; y1 := TRUE; t0_start := TRUE; t0_up := FALSE; 
    ELSIF ((x0 = FALSE) AND  (x1 = TRUE) AND  (x2 = FALSE) AND  (t0.Q = FALSE)) THEN 
        cstate58 := 6404; y0 := FALSE; y1 := FALSE; t0_start := FALSE; 
    ELSIF ((x0 = FALSE) AND  (x1 = TRUE) AND  (x2 = FALSE) AND  (t0.Q = TRUE)) THEN 
        cstate58 := 6338; y0 := FALSE; y1 := FALSE; t0_start := FALSE; 
    ELSIF ((x0 = FALSE) AND  (x1 = TRUE) AND  (x2 = TRUE) AND  (t0.Q = FALSE)) THEN 
        cstate58 := 6468; y0 := FALSE; y1 := FALSE; t0_start := TRUE; t0_up := FALSE; 
    ELSIF ((x0 = FALSE) AND  (x1 = TRUE) AND  (x2 = TRUE) AND  (t0.Q = TRUE)) THEN 
        cstate58 := 6466; y0 := FALSE; y1 := FALSE; t0_start := TRUE; t0_up := FALSE; 
    ELSIF ((x0 = TRUE) AND  (x1 = FALSE) AND  (x2 = FALSE) AND  (t0.Q = FALSE)) THEN 
        cstate58 := 5256; y0 := TRUE; y1 := FALSE; t0_start := FALSE; 
    ELSIF ((x0 = TRUE) AND  (x1 = FALSE) AND  (x2 = FALSE) AND  (t0.Q = TRUE)) THEN 
        cstate58 := 5186; y0 := TRUE; y1 := FALSE; t0_start := FALSE; 
    ELSIF ((x0 = TRUE) AND  (x1 = FALSE) AND  (x2 = TRUE) AND  (t0.Q = FALSE)) THEN 
        cstate58 := 3784; y0 := FALSE; y1 := FALSE; t0_start := TRUE; t0_up := FALSE; 
    ELSIF ((x0 = TRUE) AND  (x1 = FALSE) AND  (x2 = TRUE) AND  (t0.Q = TRUE)) THEN 
        cstate58 := 3778; y0 := FALSE; y1 := FALSE; t0_start := TRUE; t0_up := FALSE; 
    ELSIF ((x0 = TRUE) AND  (x1 = TRUE) AND  (x2 = FALSE) AND  (t0.Q = FALSE)) THEN 
        cstate58 := 4742; y0 := TRUE; y1 := FALSE; t0_start := FALSE; 
    ELSIF ((x0 = TRUE) AND  (x1 = TRUE) AND  (x2 = FALSE) AND  (t0.Q = TRUE)) THEN 
        cstate58 := 4674; y0 := TRUE; y1 := FALSE; t0_start := FALSE; 
    ELSIF ((x0 = TRUE) AND  (x1 = TRUE) AND  (x2 = TRUE) AND  (t0.Q = FALSE)) THEN 
        cstate58 := 2566; y0 := FALSE; y1 := FALSE; t0_start := TRUE; t0_up := FALSE; 
    ELSIF ((x0 = TRUE) AND  (x1 = TRUE) AND  (x2 = TRUE) AND  (t0.Q = TRUE)) THEN 
        cstate58 := 2562; y0 := FALSE; y1 := FALSE; t0_start := TRUE; t0_up := FALSE; 
    END_IF;
3778:
    IF ((x0 = FALSE) AND  (x1 = FALSE) AND  (x2 = FALSE) AND  (t0.Q = FALSE)) THEN 
        cstate58 := 7428; y0 := FALSE; y1 := FALSE; t0_start := FALSE; 
    ELSIF ((x0 = FALSE) AND  (x1 = FALSE) AND  (x2 = FALSE) AND  (t0.Q = TRUE)) THEN 
        cstate58 := 7362; y0 := FALSE; y1 := FALSE; t0_start := FALSE; 
    ELSIF ((x0 = FALSE) AND  (x1 = FALSE) AND  (x2 = TRUE) AND  (t0.Q = FALSE)) THEN 
        cstate58 := 7492; y0 := FALSE; y1 := FALSE; t0_start := FALSE; 
    ELSIF ((x0 = FALSE) AND  (x1 = FALSE) AND  (x2 = TRUE) AND  (t0.Q = TRUE)) THEN 
        cstate58 := 7554; y0 := FALSE; y1 := FALSE; t0_start := FALSE; 
    ELSIF ((x0 = FALSE) AND  (x1 = TRUE) AND  (x2 = FALSE) AND  (t0.Q = FALSE)) THEN 
        cstate58 := 6404; y0 := FALSE; y1 := FALSE; t0_start := FALSE; 
    ELSIF ((x0 = FALSE) AND  (x1 = TRUE) AND  (x2 = FALSE) AND  (t0.Q = TRUE)) THEN 
        cstate58 := 6338; y0 := FALSE; y1 := FALSE; t0_start := FALSE; 
    ELSIF ((x0 = FALSE) AND  (x1 = TRUE) AND  (x2 = TRUE) AND  (t0.Q = FALSE)) THEN 
        cstate58 := 6468; y0 := FALSE; y1 := FALSE; t0_start := FALSE; 
    ELSIF ((x0 = FALSE) AND  (x1 = TRUE) AND  (x2 = TRUE) AND  (t0.Q = TRUE)) THEN 
        cstate58 := 6530; y0 := FALSE; y1 := FALSE; t0_start := FALSE; 
    ELSIF ((x0 = TRUE) AND  (x1 = FALSE) AND  (x2 = FALSE) AND  (t0.Q = FALSE)) THEN 
        cstate58 := 3208; y0 := FALSE; y1 := FALSE; t0_start := FALSE; 
    ELSIF ((x0 = TRUE) AND  (x1 = FALSE) AND  (x2 = FALSE) AND  (t0.Q = TRUE)) THEN 
        cstate58 := 3138; y0 := FALSE; y1 := FALSE; t0_start := FALSE; 
    ELSIF ((x0 = TRUE) AND  (x1 = FALSE) AND  (x2 = TRUE) AND  (t0.Q = FALSE)) THEN 
        cstate58 := 3784; y0 := FALSE; y1 := FALSE; t0_start := FALSE; 
    ELSIF ((x0 = TRUE) AND  (x1 = FALSE) AND  (x2 = TRUE) AND  (t0.Q = TRUE)) THEN 
        cstate58 := 3842; y0 := FALSE; y1 := FALSE; t0_start := FALSE; 
    ELSIF ((x0 = TRUE) AND  (x1 = TRUE) AND  (x2 = FALSE) AND  (t0.Q = FALSE)) THEN 
        cstate58 := 2694; y0 := FALSE; y1 := FALSE; t0_start := FALSE; 
    ELSIF ((x0 = TRUE) AND  (x1 = TRUE) AND  (x2 = FALSE) AND  (t0.Q = TRUE)) THEN 
        cstate58 := 2626; y0 := FALSE; y1 := FALSE; t0_start := FALSE; 
    ELSIF ((x0 = TRUE) AND  (x1 = TRUE) AND  (x2 = TRUE) AND  (t0.Q = FALSE)) THEN 
        cstate58 := 2566; y0 := FALSE; y1 := FALSE; t0_start := FALSE; 
    ELSIF ((x0 = TRUE) AND  (x1 = TRUE) AND  (x2 = TRUE) AND  (t0.Q = TRUE)) THEN 
        cstate58 := 2498; y0 := FALSE; y1 := FALSE; t0_start := FALSE; 
    END_IF;
7390:
    IF ((x0 = FALSE) AND  (x1 = FALSE) AND  (x2 = FALSE) AND  (t0.Q = FALSE)) THEN 
        cstate58 := 7390; y0 := FALSE; y1 := TRUE; t0_start := FALSE; 
    ELSIF ((x0 = FALSE) AND  (x1 = FALSE) AND  (x2 = FALSE) AND  (t0.Q = TRUE)) THEN 
        cstate58 := 7378; y0 := FALSE; y1 := TRUE; t0_start := FALSE; 
    ELSIF ((x0 = FALSE) AND  (x1 = FALSE) AND  (x2 = TRUE) AND  (t0.Q = FALSE)) THEN 
        cstate58 := 7520; y0 := FALSE; y1 := TRUE; t0_start := TRUE; t0_up := FALSE; 
    ELSIF ((x0 = FALSE) AND  (x1 = FALSE) AND  (x2 = TRUE) AND  (t0.Q = TRUE)) THEN 
        cstate58 := 7508; y0 := FALSE; y1 := TRUE; t0_start := TRUE; t0_up := FALSE; 
    ELSIF ((x0 = FALSE) AND  (x1 = TRUE) AND  (x2 = FALSE) AND  (t0.Q = FALSE)) THEN 
        cstate58 := 6340; y0 := FALSE; y1 := FALSE; t0_start := FALSE; 
    ELSIF ((x0 = FALSE) AND  (x1 = TRUE) AND  (x2 = FALSE) AND  (t0.Q = TRUE)) THEN 
        cstate58 := 6338; y0 := FALSE; y1 := FALSE; t0_start := FALSE; 
    ELSIF ((x0 = FALSE) AND  (x1 = TRUE) AND  (x2 = TRUE) AND  (t0.Q = FALSE)) THEN 
        cstate58 := 6468; y0 := FALSE; y1 := FALSE; t0_start := TRUE; t0_up := FALSE; 
    ELSIF ((x0 = FALSE) AND  (x1 = TRUE) AND  (x2 = TRUE) AND  (t0.Q = TRUE)) THEN 
        cstate58 := 6466; y0 := FALSE; y1 := FALSE; t0_start := TRUE; t0_up := FALSE; 
    ELSIF ((x0 = TRUE) AND  (x1 = FALSE) AND  (x2 = FALSE) AND  (t0.Q = FALSE)) THEN 
        cstate58 := 5192; y0 := TRUE; y1 := FALSE; t0_start := FALSE; 
    ELSIF ((x0 = TRUE) AND  (x1 = FALSE) AND  (x2 = FALSE) AND  (t0.Q = TRUE)) THEN 
        cstate58 := 5186; y0 := TRUE; y1 := FALSE; t0_start := FALSE; 
    ELSIF ((x0 = TRUE) AND  (x1 = FALSE) AND  (x2 = TRUE) AND  (t0.Q = FALSE)) THEN 
        cstate58 := 3784; y0 := FALSE; y1 := FALSE; t0_start := TRUE; t0_up := FALSE; 
    ELSIF ((x0 = TRUE) AND  (x1 = FALSE) AND  (x2 = TRUE) AND  (t0.Q = TRUE)) THEN 
        cstate58 := 3778; y0 := FALSE; y1 := FALSE; t0_start := TRUE; t0_up := FALSE; 
    ELSIF ((x0 = TRUE) AND  (x1 = TRUE) AND  (x2 = FALSE) AND  (t0.Q = FALSE)) THEN 
        cstate58 := 4678; y0 := TRUE; y1 := FALSE; t0_start := FALSE; 
    ELSIF ((x0 = TRUE) AND  (x1 = TRUE) AND  (x2 = FALSE) AND  (t0.Q = TRUE)) THEN 
        cstate58 := 4674; y0 := TRUE; y1 := FALSE; t0_start := FALSE; 
    ELSIF ((x0 = TRUE) AND  (x1 = TRUE) AND  (x2 = TRUE) AND  (t0.Q = FALSE)) THEN 
        cstate58 := 2566; y0 := FALSE; y1 := FALSE; t0_start := TRUE; t0_up := FALSE; 
    ELSIF ((x0 = TRUE) AND  (x1 = TRUE) AND  (x2 = TRUE) AND  (t0.Q = TRUE)) THEN 
        cstate58 := 2562; y0 := FALSE; y1 := FALSE; t0_start := TRUE; t0_up := FALSE; 
    END_IF;
7500:
    IF ((x0 = FALSE) AND  (x1 = FALSE) AND  (x2 = FALSE) AND  (t0.Q = FALSE)) THEN 
        cstate58 := 7448; y0 := FALSE; y1 := TRUE; t0_start := FALSE; 
    ELSIF ((x0 = FALSE) AND  (x1 = FALSE) AND  (x2 = FALSE) AND  (t0.Q = TRUE)) THEN 
        cstate58 := 7370; y0 := FALSE; y1 := TRUE; t0_start := FALSE; 
    ELSIF ((x0 = FALSE) AND  (x1 = FALSE) AND  (x2 = TRUE) AND  (t0.Q = FALSE)) THEN 
        cstate58 := 7512; y0 := FALSE; y1 := TRUE; t0_start := FALSE; 
    ELSIF ((x0 = FALSE) AND  (x1 = FALSE) AND  (x2 = TRUE) AND  (t0.Q = TRUE)) THEN 
        cstate58 := 7562; y0 := FALSE; y1 := TRUE; t0_start := FALSE; 
    ELSIF ((x0 = FALSE) AND  (x1 = TRUE) AND  (x2 = FALSE) AND  (t0.Q = FALSE)) THEN 
        cstate58 := 6404; y0 := FALSE; y1 := FALSE; t0_start := FALSE; 
    ELSIF ((x0 = FALSE) AND  (x1 = TRUE) AND  (x2 = FALSE) AND  (t0.Q = TRUE)) THEN 
        cstate58 := 6338; y0 := FALSE; y1 := FALSE; t0_start := FALSE; 
    ELSIF ((x0 = FALSE) AND  (x1 = TRUE) AND  (x2 = TRUE) AND  (t0.Q = FALSE)) THEN 
        cstate58 := 6468; y0 := FALSE; y1 := FALSE; t0_start := FALSE; 
    ELSIF ((x0 = FALSE) AND  (x1 = TRUE) AND  (x2 = TRUE) AND  (t0.Q = TRUE)) THEN 
        cstate58 := 6530; y0 := FALSE; y1 := FALSE; t0_start := FALSE; 
    ELSIF ((x0 = TRUE) AND  (x1 = FALSE) AND  (x2 = FALSE) AND  (t0.Q = FALSE)) THEN 
        cstate58 := 5256; y0 := TRUE; y1 := FALSE; t0_start := FALSE; 
    ELSIF ((x0 = TRUE) AND  (x1 = FALSE) AND  (x2 = FALSE) AND  (t0.Q = TRUE)) THEN 
        cstate58 := 5186; y0 := TRUE; y1 := FALSE; t0_start := FALSE; 
    ELSIF ((x0 = TRUE) AND  (x1 = FALSE) AND  (x2 = TRUE) AND  (t0.Q = FALSE)) THEN 
        cstate58 := 3784; y0 := FALSE; y1 := FALSE; t0_start := FALSE; 
    ELSIF ((x0 = TRUE) AND  (x1 = FALSE) AND  (x2 = TRUE) AND  (t0.Q = TRUE)) THEN 
        cstate58 := 3842; y0 := FALSE; y1 := FALSE; t0_start := FALSE; 
    ELSIF ((x0 = TRUE) AND  (x1 = TRUE) AND  (x2 = FALSE) AND  (t0.Q = FALSE)) THEN 
        cstate58 := 4742; y0 := TRUE; y1 := FALSE; t0_start := FALSE; 
    ELSIF ((x0 = TRUE) AND  (x1 = TRUE) AND  (x2 = FALSE) AND  (t0.Q = TRUE)) THEN 
        cstate58 := 4674; y0 := TRUE; y1 := FALSE; t0_start := FALSE; 
    ELSIF ((x0 = TRUE) AND  (x1 = TRUE) AND  (x2 = TRUE) AND  (t0.Q = FALSE)) THEN 
        cstate58 := 2566; y0 := FALSE; y1 := FALSE; t0_start := FALSE; 
    ELSIF ((x0 = TRUE) AND  (x1 = TRUE) AND  (x2 = TRUE) AND  (t0.Q = TRUE)) THEN 
        cstate58 := 2498; y0 := FALSE; y1 := FALSE; t0_start := FALSE; 
    END_IF;
1348:
    IF ((x0 = FALSE) AND  (x1 = FALSE) AND  (x2 = FALSE) AND  (t0.Q = FALSE)) THEN 
        cstate58 := 1284; y0 := FALSE; y1 := FALSE; t0_start := FALSE; 
    ELSIF ((x0 = FALSE) AND  (x1 = FALSE) AND  (x2 = FALSE) AND  (t0.Q = TRUE)) THEN 
        cstate58 := 1226; y0 := FALSE; y1 := TRUE; t0_start := FALSE; 
    ELSIF ((x0 = FALSE) AND  (x1 = FALSE) AND  (x2 = TRUE) AND  (t0.Q = FALSE)) THEN 
        cstate58 := 1348; y0 := FALSE; y1 := FALSE; t0_start := FALSE; 
    ELSIF ((x0 = FALSE) AND  (x1 = FALSE) AND  (x2 = TRUE) AND  (t0.Q = TRUE)) THEN 
        cstate58 := 1418; y0 := FALSE; y1 := TRUE; t0_start := FALSE; 
    ELSIF ((x0 = FALSE) AND  (x1 = TRUE) AND  (x2 = FALSE) AND  (t0.Q = FALSE)) THEN 
        cstate58 := 1284; y0 := FALSE; y1 := FALSE; t0_start := FALSE; 
    ELSIF ((x0 = FALSE) AND  (x1 = TRUE) AND  (x2 = FALSE) AND  (t0.Q = TRUE)) THEN 
        cstate58 := 1218; y0 := FALSE; y1 := FALSE; t0_start := FALSE; 
    ELSIF ((x0 = FALSE) AND  (x1 = TRUE) AND  (x2 = TRUE) AND  (t0.Q = FALSE)) THEN 
        cstate58 := 1348; y0 := FALSE; y1 := FALSE; t0_start := FALSE; 
    ELSIF ((x0 = FALSE) AND  (x1 = TRUE) AND  (x2 = TRUE) AND  (t0.Q = TRUE)) THEN 
        cstate58 := 1410; y0 := FALSE; y1 := FALSE; t0_start := FALSE; 
    ELSIF ((x0 = TRUE) AND  (x1 = FALSE) AND  (x2 = FALSE) AND  (t0.Q = FALSE)) THEN 
        cstate58 := 5256; y0 := TRUE; y1 := FALSE; t0_start := FALSE; 
    ELSIF ((x0 = TRUE) AND  (x1 = FALSE) AND  (x2 = FALSE) AND  (t0.Q = TRUE)) THEN 
        cstate58 := 5186; y0 := TRUE; y1 := FALSE; t0_start := FALSE; 
    ELSIF ((x0 = TRUE) AND  (x1 = FALSE) AND  (x2 = TRUE) AND  (t0.Q = FALSE)) THEN 
        cstate58 := 3784; y0 := FALSE; y1 := FALSE; t0_start := FALSE; 
    ELSIF ((x0 = TRUE) AND  (x1 = FALSE) AND  (x2 = TRUE) AND  (t0.Q = TRUE)) THEN 
        cstate58 := 3842; y0 := FALSE; y1 := FALSE; t0_start := FALSE; 
    ELSIF ((x0 = TRUE) AND  (x1 = TRUE) AND  (x2 = FALSE) AND  (t0.Q = FALSE)) THEN 
        cstate58 := 4742; y0 := TRUE; y1 := FALSE; t0_start := FALSE; 
    ELSIF ((x0 = TRUE) AND  (x1 = TRUE) AND  (x2 = FALSE) AND  (t0.Q = TRUE)) THEN 
        cstate58 := 4674; y0 := TRUE; y1 := FALSE; t0_start := FALSE; 
    ELSIF ((x0 = TRUE) AND  (x1 = TRUE) AND  (x2 = TRUE) AND  (t0.Q = FALSE)) THEN 
        cstate58 := 2566; y0 := FALSE; y1 := FALSE; t0_start := FALSE; 
    ELSIF ((x0 = TRUE) AND  (x1 = TRUE) AND  (x2 = TRUE) AND  (t0.Q = TRUE)) THEN 
        cstate58 := 2498; y0 := FALSE; y1 := FALSE; t0_start := FALSE; 
    END_IF;
1346:
    IF ((x0 = FALSE) AND  (x1 = FALSE) AND  (x2 = FALSE) AND  (t0.Q = FALSE)) THEN 
        cstate58 := 1284; y0 := FALSE; y1 := FALSE; t0_start := FALSE; 
    ELSIF ((x0 = FALSE) AND  (x1 = FALSE) AND  (x2 = FALSE) AND  (t0.Q = TRUE)) THEN 
        cstate58 := 1218; y0 := FALSE; y1 := FALSE; t0_start := FALSE; 
    ELSIF ((x0 = FALSE) AND  (x1 = FALSE) AND  (x2 = TRUE) AND  (t0.Q = FALSE)) THEN 
        cstate58 := 1348; y0 := FALSE; y1 := FALSE; t0_start := FALSE; 
    ELSIF ((x0 = FALSE) AND  (x1 = FALSE) AND  (x2 = TRUE) AND  (t0.Q = TRUE)) THEN 
        cstate58 := 1410; y0 := FALSE; y1 := FALSE; t0_start := FALSE; 
    ELSIF ((x0 = FALSE) AND  (x1 = TRUE) AND  (x2 = FALSE) AND  (t0.Q = FALSE)) THEN 
        cstate58 := 1284; y0 := FALSE; y1 := FALSE; t0_start := FALSE; 
    ELSIF ((x0 = FALSE) AND  (x1 = TRUE) AND  (x2 = FALSE) AND  (t0.Q = TRUE)) THEN 
        cstate58 := 1218; y0 := FALSE; y1 := FALSE; t0_start := FALSE; 
    ELSIF ((x0 = FALSE) AND  (x1 = TRUE) AND  (x2 = TRUE) AND  (t0.Q = FALSE)) THEN 
        cstate58 := 1348; y0 := FALSE; y1 := FALSE; t0_start := FALSE; 
    ELSIF ((x0 = FALSE) AND  (x1 = TRUE) AND  (x2 = TRUE) AND  (t0.Q = TRUE)) THEN 
        cstate58 := 1410; y0 := FALSE; y1 := FALSE; t0_start := FALSE; 
    ELSIF ((x0 = TRUE) AND  (x1 = FALSE) AND  (x2 = FALSE) AND  (t0.Q = FALSE)) THEN 
        cstate58 := 5256; y0 := TRUE; y1 := FALSE; t0_start := FALSE; 
    ELSIF ((x0 = TRUE) AND  (x1 = FALSE) AND  (x2 = FALSE) AND  (t0.Q = TRUE)) THEN 
        cstate58 := 5186; y0 := TRUE; y1 := FALSE; t0_start := FALSE; 
    ELSIF ((x0 = TRUE) AND  (x1 = FALSE) AND  (x2 = TRUE) AND  (t0.Q = FALSE)) THEN 
        cstate58 := 3784; y0 := FALSE; y1 := FALSE; t0_start := FALSE; 
    ELSIF ((x0 = TRUE) AND  (x1 = FALSE) AND  (x2 = TRUE) AND  (t0.Q = TRUE)) THEN 
        cstate58 := 3842; y0 := FALSE; y1 := FALSE; t0_start := FALSE; 
    ELSIF ((x0 = TRUE) AND  (x1 = TRUE) AND  (x2 = FALSE) AND  (t0.Q = FALSE)) THEN 
        cstate58 := 4742; y0 := TRUE; y1 := FALSE; t0_start := FALSE; 
    ELSIF ((x0 = TRUE) AND  (x1 = TRUE) AND  (x2 = FALSE) AND  (t0.Q = TRUE)) THEN 
        cstate58 := 4674; y0 := TRUE; y1 := FALSE; t0_start := FALSE; 
    ELSIF ((x0 = TRUE) AND  (x1 = TRUE) AND  (x2 = TRUE) AND  (t0.Q = FALSE)) THEN 
        cstate58 := 2566; y0 := FALSE; y1 := FALSE; t0_start := FALSE; 
    ELSIF ((x0 = TRUE) AND  (x1 = TRUE) AND  (x2 = TRUE) AND  (t0.Q = TRUE)) THEN 
        cstate58 := 2498; y0 := FALSE; y1 := FALSE; t0_start := FALSE; 
    END_IF;
2502:
    IF ((x0 = FALSE) AND  (x1 = FALSE) AND  (x2 = FALSE) AND  (t0.Q = FALSE)) THEN 
        cstate58 := 6340; y0 := FALSE; y1 := FALSE; t0_start := FALSE; 
    ELSIF ((x0 = FALSE) AND  (x1 = FALSE) AND  (x2 = FALSE) AND  (t0.Q = TRUE)) THEN 
        cstate58 := 6350; y0 := FALSE; y1 := TRUE; t0_start := FALSE; 
    ELSIF ((x0 = FALSE) AND  (x1 = FALSE) AND  (x2 = TRUE) AND  (t0.Q = FALSE)) THEN 
        cstate58 := 6532; y0 := FALSE; y1 := FALSE; t0_start := FALSE; 
    ELSIF ((x0 = FALSE) AND  (x1 = FALSE) AND  (x2 = TRUE) AND  (t0.Q = TRUE)) THEN 
        cstate58 := 6542; y0 := FALSE; y1 := TRUE; t0_start := FALSE; 
    ELSIF ((x0 = FALSE) AND  (x1 = TRUE) AND  (x2 = FALSE) AND  (t0.Q = FALSE)) THEN 
        cstate58 := 6340; y0 := FALSE; y1 := FALSE; t0_start := FALSE; 
    ELSIF ((x0 = FALSE) AND  (x1 = TRUE) AND  (x2 = FALSE) AND  (t0.Q = TRUE)) THEN 
        cstate58 := 6338; y0 := FALSE; y1 := FALSE; t0_start := FALSE; 
    ELSIF ((x0 = FALSE) AND  (x1 = TRUE) AND  (x2 = TRUE) AND  (t0.Q = FALSE)) THEN 
        cstate58 := 6532; y0 := FALSE; y1 := FALSE; t0_start := FALSE; 
    ELSIF ((x0 = FALSE) AND  (x1 = TRUE) AND  (x2 = TRUE) AND  (t0.Q = TRUE)) THEN 
        cstate58 := 6530; y0 := FALSE; y1 := FALSE; t0_start := FALSE; 
    ELSIF ((x0 = TRUE) AND  (x1 = FALSE) AND  (x2 = FALSE) AND  (t0.Q = FALSE)) THEN 
        cstate58 := 2120; y0 := FALSE; y1 := FALSE; t0_start := FALSE; 
    ELSIF ((x0 = TRUE) AND  (x1 = FALSE) AND  (x2 = FALSE) AND  (t0.Q = TRUE)) THEN 
        cstate58 := 2114; y0 := FALSE; y1 := FALSE; t0_start := FALSE; 
    ELSIF ((x0 = TRUE) AND  (x1 = FALSE) AND  (x2 = TRUE) AND  (t0.Q = FALSE)) THEN 
        cstate58 := 2824; y0 := FALSE; y1 := FALSE; t0_start := FALSE; 
    ELSIF ((x0 = TRUE) AND  (x1 = FALSE) AND  (x2 = TRUE) AND  (t0.Q = TRUE)) THEN 
        cstate58 := 2818; y0 := FALSE; y1 := FALSE; t0_start := FALSE; 
    ELSIF ((x0 = TRUE) AND  (x1 = TRUE) AND  (x2 = FALSE) AND  (t0.Q = FALSE)) THEN 
        cstate58 := 2630; y0 := FALSE; y1 := FALSE; t0_start := FALSE; 
    ELSIF ((x0 = TRUE) AND  (x1 = TRUE) AND  (x2 = FALSE) AND  (t0.Q = TRUE)) THEN 
        cstate58 := 2626; y0 := FALSE; y1 := FALSE; t0_start := FALSE; 
    ELSIF ((x0 = TRUE) AND  (x1 = TRUE) AND  (x2 = TRUE) AND  (t0.Q = FALSE)) THEN 
        cstate58 := 2502; y0 := FALSE; y1 := FALSE; t0_start := FALSE; 
    ELSIF ((x0 = TRUE) AND  (x1 = TRUE) AND  (x2 = TRUE) AND  (t0.Q = TRUE)) THEN 
        cstate58 := 2498; y0 := FALSE; y1 := FALSE; t0_start := FALSE; 
    END_IF;
2120:
    IF ((x0 = FALSE) AND  (x1 = FALSE) AND  (x2 = FALSE) AND  (t0.Q = FALSE)) THEN 
        cstate58 := 6340; y0 := FALSE; y1 := FALSE; t0_start := FALSE; 
    ELSIF ((x0 = FALSE) AND  (x1 = FALSE) AND  (x2 = FALSE) AND  (t0.Q = TRUE)) THEN 
        cstate58 := 6354; y0 := FALSE; y1 := TRUE; t0_start := FALSE; 
    ELSIF ((x0 = FALSE) AND  (x1 = FALSE) AND  (x2 = TRUE) AND  (t0.Q = FALSE)) THEN 
        cstate58 := 6468; y0 := FALSE; y1 := FALSE; t0_start := TRUE; t0_up := FALSE; 
    ELSIF ((x0 = FALSE) AND  (x1 = FALSE) AND  (x2 = TRUE) AND  (t0.Q = TRUE)) THEN 
        cstate58 := 6484; y0 := FALSE; y1 := TRUE; t0_start := TRUE; t0_up := FALSE; 
    ELSIF ((x0 = FALSE) AND  (x1 = TRUE) AND  (x2 = FALSE) AND  (t0.Q = FALSE)) THEN 
        cstate58 := 6340; y0 := FALSE; y1 := FALSE; t0_start := FALSE; 
    ELSIF ((x0 = FALSE) AND  (x1 = TRUE) AND  (x2 = FALSE) AND  (t0.Q = TRUE)) THEN 
        cstate58 := 6338; y0 := FALSE; y1 := FALSE; t0_start := FALSE; 
    ELSIF ((x0 = FALSE) AND  (x1 = TRUE) AND  (x2 = TRUE) AND  (t0.Q = FALSE)) THEN 
        cstate58 := 6468; y0 := FALSE; y1 := FALSE; t0_start := TRUE; t0_up := FALSE; 
    ELSIF ((x0 = FALSE) AND  (x1 = TRUE) AND  (x2 = TRUE) AND  (t0.Q = TRUE)) THEN 
        cstate58 := 6466; y0 := FALSE; y1 := FALSE; t0_start := TRUE; t0_up := FALSE; 
    ELSIF ((x0 = TRUE) AND  (x1 = FALSE) AND  (x2 = FALSE) AND  (t0.Q = FALSE)) THEN 
        cstate58 := 2120; y0 := FALSE; y1 := FALSE; t0_start := FALSE; 
    ELSIF ((x0 = TRUE) AND  (x1 = FALSE) AND  (x2 = FALSE) AND  (t0.Q = TRUE)) THEN 
        cstate58 := 2114; y0 := FALSE; y1 := FALSE; t0_start := FALSE; 
    ELSIF ((x0 = TRUE) AND  (x1 = FALSE) AND  (x2 = TRUE) AND  (t0.Q = FALSE)) THEN 
        cstate58 := 2760; y0 := FALSE; y1 := FALSE; t0_start := TRUE; t0_up := FALSE; 
    ELSIF ((x0 = TRUE) AND  (x1 = FALSE) AND  (x2 = TRUE) AND  (t0.Q = TRUE)) THEN 
        cstate58 := 2754; y0 := FALSE; y1 := FALSE; t0_start := TRUE; t0_up := FALSE; 
    ELSIF ((x0 = TRUE) AND  (x1 = TRUE) AND  (x2 = FALSE) AND  (t0.Q = FALSE)) THEN 
        cstate58 := 2630; y0 := FALSE; y1 := FALSE; t0_start := FALSE; 
    ELSIF ((x0 = TRUE) AND  (x1 = TRUE) AND  (x2 = FALSE) AND  (t0.Q = TRUE)) THEN 
        cstate58 := 2626; y0 := FALSE; y1 := FALSE; t0_start := FALSE; 
    ELSIF ((x0 = TRUE) AND  (x1 = TRUE) AND  (x2 = TRUE) AND  (t0.Q = FALSE)) THEN 
        cstate58 := 2566; y0 := FALSE; y1 := FALSE; t0_start := TRUE; t0_up := FALSE; 
    ELSIF ((x0 = TRUE) AND  (x1 = TRUE) AND  (x2 = TRUE) AND  (t0.Q = TRUE)) THEN 
        cstate58 := 2562; y0 := FALSE; y1 := FALSE; t0_start := TRUE; t0_up := FALSE; 
    END_IF;
7582:
    IF ((x0 = FALSE) AND  (x1 = FALSE) AND  (x2 = FALSE) AND  (t0.Q = FALSE)) THEN 
        cstate58 := 7390; y0 := FALSE; y1 := TRUE; t0_start := FALSE; 
    ELSIF ((x0 = FALSE) AND  (x1 = FALSE) AND  (x2 = FALSE) AND  (t0.Q = TRUE)) THEN 
        cstate58 := 7378; y0 := FALSE; y1 := TRUE; t0_start := FALSE; 
    ELSIF ((x0 = FALSE) AND  (x1 = FALSE) AND  (x2 = TRUE) AND  (t0.Q = FALSE)) THEN 
        cstate58 := 7582; y0 := FALSE; y1 := TRUE; t0_start := FALSE; 
    ELSIF ((x0 = FALSE) AND  (x1 = FALSE) AND  (x2 = TRUE) AND  (t0.Q = TRUE)) THEN 
        cstate58 := 7570; y0 := FALSE; y1 := TRUE; t0_start := FALSE; 
    ELSIF ((x0 = FALSE) AND  (x1 = TRUE) AND  (x2 = FALSE) AND  (t0.Q = FALSE)) THEN 
        cstate58 := 6340; y0 := FALSE; y1 := FALSE; t0_start := FALSE; 
    ELSIF ((x0 = FALSE) AND  (x1 = TRUE) AND  (x2 = FALSE) AND  (t0.Q = TRUE)) THEN 
        cstate58 := 6338; y0 := FALSE; y1 := FALSE; t0_start := FALSE; 
    ELSIF ((x0 = FALSE) AND  (x1 = TRUE) AND  (x2 = TRUE) AND  (t0.Q = FALSE)) THEN 
        cstate58 := 6532; y0 := FALSE; y1 := FALSE; t0_start := FALSE; 
    ELSIF ((x0 = FALSE) AND  (x1 = TRUE) AND  (x2 = TRUE) AND  (t0.Q = TRUE)) THEN 
        cstate58 := 6530; y0 := FALSE; y1 := FALSE; t0_start := FALSE; 
    ELSIF ((x0 = TRUE) AND  (x1 = FALSE) AND  (x2 = FALSE) AND  (t0.Q = FALSE)) THEN 
        cstate58 := 5192; y0 := TRUE; y1 := FALSE; t0_start := FALSE; 
    ELSIF ((x0 = TRUE) AND  (x1 = FALSE) AND  (x2 = FALSE) AND  (t0.Q = TRUE)) THEN 
        cstate58 := 5186; y0 := TRUE; y1 := FALSE; t0_start := FALSE; 
    ELSIF ((x0 = TRUE) AND  (x1 = FALSE) AND  (x2 = TRUE) AND  (t0.Q = FALSE)) THEN 
        cstate58 := 3848; y0 := FALSE; y1 := FALSE; t0_start := FALSE; 
    ELSIF ((x0 = TRUE) AND  (x1 = FALSE) AND  (x2 = TRUE) AND  (t0.Q = TRUE)) THEN 
        cstate58 := 3842; y0 := FALSE; y1 := FALSE; t0_start := FALSE; 
    ELSIF ((x0 = TRUE) AND  (x1 = TRUE) AND  (x2 = FALSE) AND  (t0.Q = FALSE)) THEN 
        cstate58 := 4678; y0 := TRUE; y1 := FALSE; t0_start := FALSE; 
    ELSIF ((x0 = TRUE) AND  (x1 = TRUE) AND  (x2 = FALSE) AND  (t0.Q = TRUE)) THEN 
        cstate58 := 4674; y0 := TRUE; y1 := FALSE; t0_start := FALSE; 
    ELSIF ((x0 = TRUE) AND  (x1 = TRUE) AND  (x2 = TRUE) AND  (t0.Q = FALSE)) THEN 
        cstate58 := 2502; y0 := FALSE; y1 := FALSE; t0_start := FALSE; 
    ELSIF ((x0 = TRUE) AND  (x1 = TRUE) AND  (x2 = TRUE) AND  (t0.Q = TRUE)) THEN 
        cstate58 := 2498; y0 := FALSE; y1 := FALSE; t0_start := FALSE; 
    END_IF;
4742:
    IF ((x0 = FALSE) AND  ( TRUE ) AND  (x2 = FALSE) AND  (t0.Q = FALSE)) THEN 
        cstate58 := 8452; y0 := TRUE; y1 := FALSE; t0_start := FALSE; 
    ELSIF ((x0 = FALSE) AND  ( TRUE ) AND  (x2 = FALSE) AND  (t0.Q = TRUE)) THEN 
        cstate58 := 8386; y0 := TRUE; y1 := FALSE; t0_start := FALSE; 
    ELSIF ((x0 = FALSE) AND  (x1 = FALSE) AND  (x2 = TRUE) AND  (t0.Q = FALSE)) THEN 
        cstate58 := 6468; y0 := FALSE; y1 := FALSE; t0_start := TRUE; t0_up := FALSE; 
    ELSIF ((x0 = FALSE) AND  (x1 = FALSE) AND  (x2 = TRUE) AND  (t0.Q = TRUE)) THEN 
        cstate58 := 6480; y0 := FALSE; y1 := TRUE; t0_start := TRUE; t0_up := FALSE; 
    ELSIF ((x0 = FALSE) AND  (x1 = TRUE) AND  (x2 = TRUE) AND  (t0.Q = FALSE)) THEN 
        cstate58 := 6468; y0 := FALSE; y1 := FALSE; t0_start := TRUE; t0_up := FALSE; 
    ELSIF ((x0 = FALSE) AND  (x1 = TRUE) AND  (x2 = TRUE) AND  (t0.Q = TRUE)) THEN 
        cstate58 := 6466; y0 := FALSE; y1 := FALSE; t0_start := TRUE; t0_up := FALSE; 
    ELSIF ((x0 = TRUE) AND  (x1 = FALSE) AND  (x2 = FALSE) AND  (t0.Q = FALSE)) THEN 
        cstate58 := 4232; y0 := TRUE; y1 := FALSE; t0_start := FALSE; 
    ELSIF ((x0 = TRUE) AND  (x1 = FALSE) AND  (x2 = FALSE) AND  (t0.Q = TRUE)) THEN 
        cstate58 := 4162; y0 := TRUE; y1 := FALSE; t0_start := FALSE; 
    ELSIF ((x0 = TRUE) AND  (x1 = FALSE) AND  (x2 = TRUE) AND  (t0.Q = FALSE)) THEN 
        cstate58 := 2760; y0 := FALSE; y1 := FALSE; t0_start := TRUE; t0_up := FALSE; 
    ELSIF ((x0 = TRUE) AND  (x1 = FALSE) AND  (x2 = TRUE) AND  (t0.Q = TRUE)) THEN 
        cstate58 := 2754; y0 := FALSE; y1 := FALSE; t0_start := TRUE; t0_up := FALSE; 
    ELSIF ((x0 = TRUE) AND  (x1 = TRUE) AND  (x2 = FALSE) AND  (t0.Q = FALSE)) THEN 
        cstate58 := 4742; y0 := TRUE; y1 := FALSE; t0_start := FALSE; 
    ELSIF ((x0 = TRUE) AND  (x1 = TRUE) AND  (x2 = FALSE) AND  (t0.Q = TRUE)) THEN 
        cstate58 := 4674; y0 := TRUE; y1 := FALSE; t0_start := FALSE; 
    ELSIF ((x0 = TRUE) AND  (x1 = TRUE) AND  (x2 = TRUE) AND  (t0.Q = FALSE)) THEN 
        cstate58 := 2566; y0 := FALSE; y1 := FALSE; t0_start := TRUE; t0_up := FALSE; 
    ELSIF ((x0 = TRUE) AND  (x1 = TRUE) AND  (x2 = TRUE) AND  (t0.Q = TRUE)) THEN 
        cstate58 := 2562; y0 := FALSE; y1 := FALSE; t0_start := TRUE; t0_up := FALSE; 
    END_IF;
7508:
    IF ((x0 = FALSE) AND  (x1 = FALSE) AND  (x2 = FALSE) AND  (t0.Q = FALSE)) THEN 
        cstate58 := 7456; y0 := FALSE; y1 := TRUE; t0_start := FALSE; 
    ELSIF ((x0 = FALSE) AND  (x1 = FALSE) AND  (x2 = FALSE) AND  (t0.Q = TRUE)) THEN 
        cstate58 := 7378; y0 := FALSE; y1 := TRUE; t0_start := FALSE; 
    ELSIF ((x0 = FALSE) AND  (x1 = FALSE) AND  (x2 = TRUE) AND  (t0.Q = FALSE)) THEN 
        cstate58 := 7520; y0 := FALSE; y1 := TRUE; t0_start := FALSE; 
    ELSIF ((x0 = FALSE) AND  (x1 = FALSE) AND  (x2 = TRUE) AND  (t0.Q = TRUE)) THEN 
        cstate58 := 7570; y0 := FALSE; y1 := TRUE; t0_start := FALSE; 
    ELSIF ((x0 = FALSE) AND  (x1 = TRUE) AND  (x2 = FALSE) AND  (t0.Q = FALSE)) THEN 
        cstate58 := 6404; y0 := FALSE; y1 := FALSE; t0_start := FALSE; 
    ELSIF ((x0 = FALSE) AND  (x1 = TRUE) AND  (x2 = FALSE) AND  (t0.Q = TRUE)) THEN 
        cstate58 := 6338; y0 := FALSE; y1 := FALSE; t0_start := FALSE; 
    ELSIF ((x0 = FALSE) AND  (x1 = TRUE) AND  (x2 = TRUE) AND  (t0.Q = FALSE)) THEN 
        cstate58 := 6468; y0 := FALSE; y1 := FALSE; t0_start := FALSE; 
    ELSIF ((x0 = FALSE) AND  (x1 = TRUE) AND  (x2 = TRUE) AND  (t0.Q = TRUE)) THEN 
        cstate58 := 6530; y0 := FALSE; y1 := FALSE; t0_start := FALSE; 
    ELSIF ((x0 = TRUE) AND  (x1 = FALSE) AND  (x2 = FALSE) AND  (t0.Q = FALSE)) THEN 
        cstate58 := 5256; y0 := TRUE; y1 := FALSE; t0_start := FALSE; 
    ELSIF ((x0 = TRUE) AND  (x1 = FALSE) AND  (x2 = FALSE) AND  (t0.Q = TRUE)) THEN 
        cstate58 := 5186; y0 := TRUE; y1 := FALSE; t0_start := FALSE; 
    ELSIF ((x0 = TRUE) AND  (x1 = FALSE) AND  (x2 = TRUE) AND  (t0.Q = FALSE)) THEN 
        cstate58 := 3784; y0 := FALSE; y1 := FALSE; t0_start := FALSE; 
    ELSIF ((x0 = TRUE) AND  (x1 = FALSE) AND  (x2 = TRUE) AND  (t0.Q = TRUE)) THEN 
        cstate58 := 3842; y0 := FALSE; y1 := FALSE; t0_start := FALSE; 
    ELSIF ((x0 = TRUE) AND  (x1 = TRUE) AND  (x2 = FALSE) AND  (t0.Q = FALSE)) THEN 
        cstate58 := 4742; y0 := TRUE; y1 := FALSE; t0_start := FALSE; 
    ELSIF ((x0 = TRUE) AND  (x1 = TRUE) AND  (x2 = FALSE) AND  (t0.Q = TRUE)) THEN 
        cstate58 := 4674; y0 := TRUE; y1 := FALSE; t0_start := FALSE; 
    ELSIF ((x0 = TRUE) AND  (x1 = TRUE) AND  (x2 = TRUE) AND  (t0.Q = FALSE)) THEN 
        cstate58 := 2566; y0 := FALSE; y1 := FALSE; t0_start := FALSE; 
    ELSIF ((x0 = TRUE) AND  (x1 = TRUE) AND  (x2 = TRUE) AND  (t0.Q = TRUE)) THEN 
        cstate58 := 2498; y0 := FALSE; y1 := FALSE; t0_start := FALSE; 
    END_IF;
7382:
    IF ((x0 = FALSE) AND  (x1 = FALSE) AND  (x2 = FALSE) AND  (t0.Q = FALSE)) THEN 
        cstate58 := 7382; y0 := FALSE; y1 := TRUE; t0_start := FALSE; 
    ELSIF ((x0 = FALSE) AND  (x1 = FALSE) AND  (x2 = FALSE) AND  (t0.Q = TRUE)) THEN 
        cstate58 := 7370; y0 := FALSE; y1 := TRUE; t0_start := FALSE; 
    ELSIF ((x0 = FALSE) AND  (x1 = FALSE) AND  (x2 = TRUE) AND  (t0.Q = FALSE)) THEN 
        cstate58 := 7512; y0 := FALSE; y1 := TRUE; t0_start := TRUE; t0_up := FALSE; 
    ELSIF ((x0 = FALSE) AND  (x1 = FALSE) AND  (x2 = TRUE) AND  (t0.Q = TRUE)) THEN 
        cstate58 := 7500; y0 := FALSE; y1 := TRUE; t0_start := TRUE; t0_up := FALSE; 
    ELSIF ((x0 = FALSE) AND  (x1 = TRUE) AND  (x2 = FALSE) AND  (t0.Q = FALSE)) THEN 
        cstate58 := 6340; y0 := FALSE; y1 := FALSE; t0_start := FALSE; 
    ELSIF ((x0 = FALSE) AND  (x1 = TRUE) AND  (x2 = FALSE) AND  (t0.Q = TRUE)) THEN 
        cstate58 := 6338; y0 := FALSE; y1 := FALSE; t0_start := FALSE; 
    ELSIF ((x0 = FALSE) AND  (x1 = TRUE) AND  (x2 = TRUE) AND  (t0.Q = FALSE)) THEN 
        cstate58 := 6468; y0 := FALSE; y1 := FALSE; t0_start := TRUE; t0_up := FALSE; 
    ELSIF ((x0 = FALSE) AND  (x1 = TRUE) AND  (x2 = TRUE) AND  (t0.Q = TRUE)) THEN 
        cstate58 := 6466; y0 := FALSE; y1 := FALSE; t0_start := TRUE; t0_up := FALSE; 
    ELSIF ((x0 = TRUE) AND  (x1 = FALSE) AND  (x2 = FALSE) AND  (t0.Q = FALSE)) THEN 
        cstate58 := 5192; y0 := TRUE; y1 := FALSE; t0_start := FALSE; 
    ELSIF ((x0 = TRUE) AND  (x1 = FALSE) AND  (x2 = FALSE) AND  (t0.Q = TRUE)) THEN 
        cstate58 := 5186; y0 := TRUE; y1 := FALSE; t0_start := FALSE; 
    ELSIF ((x0 = TRUE) AND  (x1 = FALSE) AND  (x2 = TRUE) AND  (t0.Q = FALSE)) THEN 
        cstate58 := 3784; y0 := FALSE; y1 := FALSE; t0_start := TRUE; t0_up := FALSE; 
    ELSIF ((x0 = TRUE) AND  (x1 = FALSE) AND  (x2 = TRUE) AND  (t0.Q = TRUE)) THEN 
        cstate58 := 3778; y0 := FALSE; y1 := FALSE; t0_start := TRUE; t0_up := FALSE; 
    ELSIF ((x0 = TRUE) AND  (x1 = TRUE) AND  (x2 = FALSE) AND  (t0.Q = FALSE)) THEN 
        cstate58 := 4678; y0 := TRUE; y1 := FALSE; t0_start := FALSE; 
    ELSIF ((x0 = TRUE) AND  (x1 = TRUE) AND  (x2 = FALSE) AND  (t0.Q = TRUE)) THEN 
        cstate58 := 4674; y0 := TRUE; y1 := FALSE; t0_start := FALSE; 
    ELSIF ((x0 = TRUE) AND  (x1 = TRUE) AND  (x2 = TRUE) AND  (t0.Q = FALSE)) THEN 
        cstate58 := 2566; y0 := FALSE; y1 := FALSE; t0_start := TRUE; t0_up := FALSE; 
    ELSIF ((x0 = TRUE) AND  (x1 = TRUE) AND  (x2 = TRUE) AND  (t0.Q = TRUE)) THEN 
        cstate58 := 2562; y0 := FALSE; y1 := FALSE; t0_start := TRUE; t0_up := FALSE; 
    END_IF;
3784:
    IF ((x0 = FALSE) AND  (x1 = FALSE) AND  (x2 = FALSE) AND  (t0.Q = FALSE)) THEN 
        cstate58 := 7428; y0 := FALSE; y1 := FALSE; t0_start := FALSE; 
    ELSIF ((x0 = FALSE) AND  (x1 = FALSE) AND  (x2 = FALSE) AND  (t0.Q = TRUE)) THEN 
        cstate58 := 7378; y0 := FALSE; y1 := TRUE; t0_start := FALSE; 
    ELSIF ((x0 = FALSE) AND  (x1 = FALSE) AND  (x2 = TRUE) AND  (t0.Q = FALSE)) THEN 
        cstate58 := 7492; y0 := FALSE; y1 := FALSE; t0_start := FALSE; 
    ELSIF ((x0 = FALSE) AND  (x1 = FALSE) AND  (x2 = TRUE) AND  (t0.Q = TRUE)) THEN 
        cstate58 := 7570; y0 := FALSE; y1 := TRUE; t0_start := FALSE; 
    ELSIF ((x0 = FALSE) AND  (x1 = TRUE) AND  (x2 = FALSE) AND  (t0.Q = FALSE)) THEN 
        cstate58 := 6404; y0 := FALSE; y1 := FALSE; t0_start := FALSE; 
    ELSIF ((x0 = FALSE) AND  (x1 = TRUE) AND  (x2 = FALSE) AND  (t0.Q = TRUE)) THEN 
        cstate58 := 6338; y0 := FALSE; y1 := FALSE; t0_start := FALSE; 
    ELSIF ((x0 = FALSE) AND  (x1 = TRUE) AND  (x2 = TRUE) AND  (t0.Q = FALSE)) THEN 
        cstate58 := 6468; y0 := FALSE; y1 := FALSE; t0_start := FALSE; 
    ELSIF ((x0 = FALSE) AND  (x1 = TRUE) AND  (x2 = TRUE) AND  (t0.Q = TRUE)) THEN 
        cstate58 := 6530; y0 := FALSE; y1 := FALSE; t0_start := FALSE; 
    ELSIF ((x0 = TRUE) AND  (x1 = FALSE) AND  (x2 = FALSE) AND  (t0.Q = FALSE)) THEN 
        cstate58 := 3208; y0 := FALSE; y1 := FALSE; t0_start := FALSE; 
    ELSIF ((x0 = TRUE) AND  (x1 = FALSE) AND  (x2 = FALSE) AND  (t0.Q = TRUE)) THEN 
        cstate58 := 3138; y0 := FALSE; y1 := FALSE; t0_start := FALSE; 
    ELSIF ((x0 = TRUE) AND  (x1 = FALSE) AND  (x2 = TRUE) AND  (t0.Q = FALSE)) THEN 
        cstate58 := 3784; y0 := FALSE; y1 := FALSE; t0_start := FALSE; 
    ELSIF ((x0 = TRUE) AND  (x1 = FALSE) AND  (x2 = TRUE) AND  (t0.Q = TRUE)) THEN 
        cstate58 := 3842; y0 := FALSE; y1 := FALSE; t0_start := FALSE; 
    ELSIF ((x0 = TRUE) AND  (x1 = TRUE) AND  (x2 = FALSE) AND  (t0.Q = FALSE)) THEN 
        cstate58 := 2694; y0 := FALSE; y1 := FALSE; t0_start := FALSE; 
    ELSIF ((x0 = TRUE) AND  (x1 = TRUE) AND  (x2 = FALSE) AND  (t0.Q = TRUE)) THEN 
        cstate58 := 2626; y0 := FALSE; y1 := FALSE; t0_start := FALSE; 
    ELSIF ((x0 = TRUE) AND  (x1 = TRUE) AND  (x2 = TRUE) AND  (t0.Q = FALSE)) THEN 
        cstate58 := 2566; y0 := FALSE; y1 := FALSE; t0_start := FALSE; 
    ELSIF ((x0 = TRUE) AND  (x1 = TRUE) AND  (x2 = TRUE) AND  (t0.Q = TRUE)) THEN 
        cstate58 := 2498; y0 := FALSE; y1 := FALSE; t0_start := FALSE; 
    END_IF;
7512:
    IF ((x0 = FALSE) AND  (x1 = FALSE) AND  (x2 = FALSE) AND  (t0.Q = FALSE)) THEN 
        cstate58 := 7448; y0 := FALSE; y1 := TRUE; t0_start := FALSE; 
    ELSIF ((x0 = FALSE) AND  (x1 = FALSE) AND  (x2 = FALSE) AND  (t0.Q = TRUE)) THEN 
        cstate58 := 7370; y0 := FALSE; y1 := TRUE; t0_start := FALSE; 
    ELSIF ((x0 = FALSE) AND  (x1 = FALSE) AND  (x2 = TRUE) AND  (t0.Q = FALSE)) THEN 
        cstate58 := 7512; y0 := FALSE; y1 := TRUE; t0_start := FALSE; 
    ELSIF ((x0 = FALSE) AND  (x1 = FALSE) AND  (x2 = TRUE) AND  (t0.Q = TRUE)) THEN 
        cstate58 := 7562; y0 := FALSE; y1 := TRUE; t0_start := FALSE; 
    ELSIF ((x0 = FALSE) AND  (x1 = TRUE) AND  (x2 = FALSE) AND  (t0.Q = FALSE)) THEN 
        cstate58 := 6404; y0 := FALSE; y1 := FALSE; t0_start := FALSE; 
    ELSIF ((x0 = FALSE) AND  (x1 = TRUE) AND  (x2 = FALSE) AND  (t0.Q = TRUE)) THEN 
        cstate58 := 6338; y0 := FALSE; y1 := FALSE; t0_start := FALSE; 
    ELSIF ((x0 = FALSE) AND  (x1 = TRUE) AND  (x2 = TRUE) AND  (t0.Q = FALSE)) THEN 
        cstate58 := 6468; y0 := FALSE; y1 := FALSE; t0_start := FALSE; 
    ELSIF ((x0 = FALSE) AND  (x1 = TRUE) AND  (x2 = TRUE) AND  (t0.Q = TRUE)) THEN 
        cstate58 := 6530; y0 := FALSE; y1 := FALSE; t0_start := FALSE; 
    ELSIF ((x0 = TRUE) AND  (x1 = FALSE) AND  (x2 = FALSE) AND  (t0.Q = FALSE)) THEN 
        cstate58 := 5256; y0 := TRUE; y1 := FALSE; t0_start := FALSE; 
    ELSIF ((x0 = TRUE) AND  (x1 = FALSE) AND  (x2 = FALSE) AND  (t0.Q = TRUE)) THEN 
        cstate58 := 5186; y0 := TRUE; y1 := FALSE; t0_start := FALSE; 
    ELSIF ((x0 = TRUE) AND  (x1 = FALSE) AND  (x2 = TRUE) AND  (t0.Q = FALSE)) THEN 
        cstate58 := 3784; y0 := FALSE; y1 := FALSE; t0_start := FALSE; 
    ELSIF ((x0 = TRUE) AND  (x1 = FALSE) AND  (x2 = TRUE) AND  (t0.Q = TRUE)) THEN 
        cstate58 := 3842; y0 := FALSE; y1 := FALSE; t0_start := FALSE; 
    ELSIF ((x0 = TRUE) AND  (x1 = TRUE) AND  (x2 = FALSE) AND  (t0.Q = FALSE)) THEN 
        cstate58 := 4742; y0 := TRUE; y1 := FALSE; t0_start := FALSE; 
    ELSIF ((x0 = TRUE) AND  (x1 = TRUE) AND  (x2 = FALSE) AND  (t0.Q = TRUE)) THEN 
        cstate58 := 4674; y0 := TRUE; y1 := FALSE; t0_start := FALSE; 
    ELSIF ((x0 = TRUE) AND  (x1 = TRUE) AND  (x2 = TRUE) AND  (t0.Q = FALSE)) THEN 
        cstate58 := 2566; y0 := FALSE; y1 := FALSE; t0_start := FALSE; 
    ELSIF ((x0 = TRUE) AND  (x1 = TRUE) AND  (x2 = TRUE) AND  (t0.Q = TRUE)) THEN 
        cstate58 := 2498; y0 := FALSE; y1 := FALSE; t0_start := FALSE; 
    END_IF;
8452:
    IF ((x0 = FALSE) AND  ( TRUE ) AND  (x2 = FALSE) AND  (t0.Q = FALSE)) THEN 
        cstate58 := 8452; y0 := TRUE; y1 := FALSE; t0_start := FALSE; 
    ELSIF ((x0 = FALSE) AND  ( TRUE ) AND  (x2 = FALSE) AND  (t0.Q = TRUE)) THEN 
        cstate58 := 8386; y0 := TRUE; y1 := FALSE; t0_start := FALSE; 
    ELSIF ((x0 = FALSE) AND  (x1 = FALSE) AND  (x2 = TRUE) AND  (t0.Q = FALSE)) THEN 
        cstate58 := 6468; y0 := FALSE; y1 := FALSE; t0_start := TRUE; t0_up := FALSE; 
    ELSIF ((x0 = FALSE) AND  (x1 = FALSE) AND  (x2 = TRUE) AND  (t0.Q = TRUE)) THEN 
        cstate58 := 6476; y0 := FALSE; y1 := TRUE; t0_start := TRUE; t0_up := FALSE; 
    ELSIF ((x0 = FALSE) AND  (x1 = TRUE) AND  (x2 = TRUE) AND  (t0.Q = FALSE)) THEN 
        cstate58 := 6468; y0 := FALSE; y1 := FALSE; t0_start := TRUE; t0_up := FALSE; 
    ELSIF ((x0 = FALSE) AND  (x1 = TRUE) AND  (x2 = TRUE) AND  (t0.Q = TRUE)) THEN 
        cstate58 := 6466; y0 := FALSE; y1 := FALSE; t0_start := TRUE; t0_up := FALSE; 
    ELSIF ((x0 = TRUE) AND  (x1 = FALSE) AND  (x2 = FALSE) AND  (t0.Q = FALSE)) THEN 
        cstate58 := 4232; y0 := TRUE; y1 := FALSE; t0_start := FALSE; 
    ELSIF ((x0 = TRUE) AND  (x1 = FALSE) AND  (x2 = FALSE) AND  (t0.Q = TRUE)) THEN 
        cstate58 := 4162; y0 := TRUE; y1 := FALSE; t0_start := FALSE; 
    ELSIF ((x0 = TRUE) AND  (x1 = FALSE) AND  (x2 = TRUE) AND  (t0.Q = FALSE)) THEN 
        cstate58 := 2760; y0 := FALSE; y1 := FALSE; t0_start := TRUE; t0_up := FALSE; 
    ELSIF ((x0 = TRUE) AND  (x1 = FALSE) AND  (x2 = TRUE) AND  (t0.Q = TRUE)) THEN 
        cstate58 := 2754; y0 := FALSE; y1 := FALSE; t0_start := TRUE; t0_up := FALSE; 
    ELSIF ((x0 = TRUE) AND  (x1 = TRUE) AND  (x2 = FALSE) AND  (t0.Q = FALSE)) THEN 
        cstate58 := 4742; y0 := TRUE; y1 := FALSE; t0_start := FALSE; 
    ELSIF ((x0 = TRUE) AND  (x1 = TRUE) AND  (x2 = FALSE) AND  (t0.Q = TRUE)) THEN 
        cstate58 := 4674; y0 := TRUE; y1 := FALSE; t0_start := FALSE; 
    ELSIF ((x0 = TRUE) AND  (x1 = TRUE) AND  (x2 = TRUE) AND  (t0.Q = FALSE)) THEN 
        cstate58 := 2566; y0 := FALSE; y1 := FALSE; t0_start := TRUE; t0_up := FALSE; 
    ELSIF ((x0 = TRUE) AND  (x1 = TRUE) AND  (x2 = TRUE) AND  (t0.Q = TRUE)) THEN 
        cstate58 := 2562; y0 := FALSE; y1 := FALSE; t0_start := TRUE; t0_up := FALSE; 
    END_IF;
1238:
    IF ((x0 = FALSE) AND  (x1 = FALSE) AND  (x2 = FALSE) AND  (t0.Q = FALSE)) THEN 
        cstate58 := 1238; y0 := FALSE; y1 := TRUE; t0_start := FALSE; 
    ELSIF ((x0 = FALSE) AND  (x1 = FALSE) AND  (x2 = FALSE) AND  (t0.Q = TRUE)) THEN 
        cstate58 := 1226; y0 := FALSE; y1 := TRUE; t0_start := FALSE; 
    ELSIF ((x0 = FALSE) AND  (x1 = FALSE) AND  (x2 = TRUE) AND  (t0.Q = FALSE)) THEN 
        cstate58 := 1368; y0 := FALSE; y1 := TRUE; t0_start := TRUE; t0_up := FALSE; 
    ELSIF ((x0 = FALSE) AND  (x1 = FALSE) AND  (x2 = TRUE) AND  (t0.Q = TRUE)) THEN 
        cstate58 := 1356; y0 := FALSE; y1 := TRUE; t0_start := TRUE; t0_up := FALSE; 
    ELSIF ((x0 = FALSE) AND  (x1 = TRUE) AND  (x2 = FALSE) AND  (t0.Q = FALSE)) THEN 
        cstate58 := 1220; y0 := FALSE; y1 := FALSE; t0_start := FALSE; 
    ELSIF ((x0 = FALSE) AND  (x1 = TRUE) AND  (x2 = FALSE) AND  (t0.Q = TRUE)) THEN 
        cstate58 := 1218; y0 := FALSE; y1 := FALSE; t0_start := FALSE; 
    ELSIF ((x0 = FALSE) AND  (x1 = TRUE) AND  (x2 = TRUE) AND  (t0.Q = FALSE)) THEN 
        cstate58 := 1348; y0 := FALSE; y1 := FALSE; t0_start := TRUE; t0_up := FALSE; 
    ELSIF ((x0 = FALSE) AND  (x1 = TRUE) AND  (x2 = TRUE) AND  (t0.Q = TRUE)) THEN 
        cstate58 := 1346; y0 := FALSE; y1 := FALSE; t0_start := TRUE; t0_up := FALSE; 
    ELSIF ((x0 = TRUE) AND  (x1 = FALSE) AND  (x2 = FALSE) AND  (t0.Q = FALSE)) THEN 
        cstate58 := 5192; y0 := TRUE; y1 := FALSE; t0_start := FALSE; 
    ELSIF ((x0 = TRUE) AND  (x1 = FALSE) AND  (x2 = FALSE) AND  (t0.Q = TRUE)) THEN 
        cstate58 := 5186; y0 := TRUE; y1 := FALSE; t0_start := FALSE; 
    ELSIF ((x0 = TRUE) AND  (x1 = FALSE) AND  (x2 = TRUE) AND  (t0.Q = FALSE)) THEN 
        cstate58 := 3784; y0 := FALSE; y1 := FALSE; t0_start := TRUE; t0_up := FALSE; 
    ELSIF ((x0 = TRUE) AND  (x1 = FALSE) AND  (x2 = TRUE) AND  (t0.Q = TRUE)) THEN 
        cstate58 := 3778; y0 := FALSE; y1 := FALSE; t0_start := TRUE; t0_up := FALSE; 
    ELSIF ((x0 = TRUE) AND  (x1 = TRUE) AND  (x2 = FALSE) AND  (t0.Q = FALSE)) THEN 
        cstate58 := 4678; y0 := TRUE; y1 := FALSE; t0_start := FALSE; 
    ELSIF ((x0 = TRUE) AND  (x1 = TRUE) AND  (x2 = FALSE) AND  (t0.Q = TRUE)) THEN 
        cstate58 := 4674; y0 := TRUE; y1 := FALSE; t0_start := FALSE; 
    ELSIF ((x0 = TRUE) AND  (x1 = TRUE) AND  (x2 = TRUE) AND  (t0.Q = FALSE)) THEN 
        cstate58 := 2566; y0 := FALSE; y1 := FALSE; t0_start := TRUE; t0_up := FALSE; 
    ELSIF ((x0 = TRUE) AND  (x1 = TRUE) AND  (x2 = TRUE) AND  (t0.Q = TRUE)) THEN 
        cstate58 := 2562; y0 := FALSE; y1 := FALSE; t0_start := TRUE; t0_up := FALSE; 
    END_IF;
4162:
    IF ((x0 = FALSE) AND  ( TRUE ) AND  (x2 = FALSE) AND  (t0.Q = FALSE)) THEN 
        cstate58 := 8388; y0 := TRUE; y1 := FALSE; t0_start := FALSE; 
    ELSIF ((x0 = FALSE) AND  ( TRUE ) AND  (x2 = FALSE) AND  (t0.Q = TRUE)) THEN 
        cstate58 := 8386; y0 := TRUE; y1 := FALSE; t0_start := FALSE; 
    ELSIF ((x0 = FALSE) AND  (x1 = FALSE) AND  (x2 = TRUE) AND  (t0.Q = FALSE)) THEN 
        cstate58 := 6468; y0 := FALSE; y1 := FALSE; t0_start := TRUE; t0_up := FALSE; 
    ELSIF ((x0 = FALSE) AND  (x1 = FALSE) AND  (x2 = TRUE) AND  (t0.Q = TRUE)) THEN 
        cstate58 := 6466; y0 := FALSE; y1 := FALSE; t0_start := TRUE; t0_up := FALSE; 
    ELSIF ((x0 = FALSE) AND  (x1 = TRUE) AND  (x2 = TRUE) AND  (t0.Q = FALSE)) THEN 
        cstate58 := 6468; y0 := FALSE; y1 := FALSE; t0_start := TRUE; t0_up := FALSE; 
    ELSIF ((x0 = FALSE) AND  (x1 = TRUE) AND  (x2 = TRUE) AND  (t0.Q = TRUE)) THEN 
        cstate58 := 6466; y0 := FALSE; y1 := FALSE; t0_start := TRUE; t0_up := FALSE; 
    ELSIF ((x0 = TRUE) AND  (x1 = FALSE) AND  (x2 = FALSE) AND  (t0.Q = FALSE)) THEN 
        cstate58 := 4168; y0 := TRUE; y1 := FALSE; t0_start := FALSE; 
    ELSIF ((x0 = TRUE) AND  (x1 = FALSE) AND  (x2 = FALSE) AND  (t0.Q = TRUE)) THEN 
        cstate58 := 4162; y0 := TRUE; y1 := FALSE; t0_start := FALSE; 
    ELSIF ((x0 = TRUE) AND  (x1 = FALSE) AND  (x2 = TRUE) AND  (t0.Q = FALSE)) THEN 
        cstate58 := 2760; y0 := FALSE; y1 := FALSE; t0_start := TRUE; t0_up := FALSE; 
    ELSIF ((x0 = TRUE) AND  (x1 = FALSE) AND  (x2 = TRUE) AND  (t0.Q = TRUE)) THEN 
        cstate58 := 2754; y0 := FALSE; y1 := FALSE; t0_start := TRUE; t0_up := FALSE; 
    ELSIF ((x0 = TRUE) AND  (x1 = TRUE) AND  (x2 = FALSE) AND  (t0.Q = FALSE)) THEN 
        cstate58 := 4678; y0 := TRUE; y1 := FALSE; t0_start := FALSE; 
    ELSIF ((x0 = TRUE) AND  (x1 = TRUE) AND  (x2 = FALSE) AND  (t0.Q = TRUE)) THEN 
        cstate58 := 4674; y0 := TRUE; y1 := FALSE; t0_start := FALSE; 
    ELSIF ((x0 = TRUE) AND  (x1 = TRUE) AND  (x2 = TRUE) AND  (t0.Q = FALSE)) THEN 
        cstate58 := 2566; y0 := FALSE; y1 := FALSE; t0_start := TRUE; t0_up := FALSE; 
    ELSIF ((x0 = TRUE) AND  (x1 = TRUE) AND  (x2 = TRUE) AND  (t0.Q = TRUE)) THEN 
        cstate58 := 2562; y0 := FALSE; y1 := FALSE; t0_start := TRUE; t0_up := FALSE; 
    END_IF;
2114:
    IF ((x0 = FALSE) AND  (x1 = FALSE) AND  (x2 = FALSE) AND  (t0.Q = FALSE)) THEN 
        cstate58 := 6340; y0 := FALSE; y1 := FALSE; t0_start := FALSE; 
    ELSIF ((x0 = FALSE) AND  (x1 = FALSE) AND  (x2 = FALSE) AND  (t0.Q = TRUE)) THEN 
        cstate58 := 6338; y0 := FALSE; y1 := FALSE; t0_start := FALSE; 
    ELSIF ((x0 = FALSE) AND  (x1 = FALSE) AND  (x2 = TRUE) AND  (t0.Q = FALSE)) THEN 
        cstate58 := 6468; y0 := FALSE; y1 := FALSE; t0_start := TRUE; t0_up := FALSE; 
    ELSIF ((x0 = FALSE) AND  (x1 = FALSE) AND  (x2 = TRUE) AND  (t0.Q = TRUE)) THEN 
        cstate58 := 6466; y0 := FALSE; y1 := FALSE; t0_start := TRUE; t0_up := FALSE; 
    ELSIF ((x0 = FALSE) AND  (x1 = TRUE) AND  (x2 = FALSE) AND  (t0.Q = FALSE)) THEN 
        cstate58 := 6340; y0 := FALSE; y1 := FALSE; t0_start := FALSE; 
    ELSIF ((x0 = FALSE) AND  (x1 = TRUE) AND  (x2 = FALSE) AND  (t0.Q = TRUE)) THEN 
        cstate58 := 6338; y0 := FALSE; y1 := FALSE; t0_start := FALSE; 
    ELSIF ((x0 = FALSE) AND  (x1 = TRUE) AND  (x2 = TRUE) AND  (t0.Q = FALSE)) THEN 
        cstate58 := 6468; y0 := FALSE; y1 := FALSE; t0_start := TRUE; t0_up := FALSE; 
    ELSIF ((x0 = FALSE) AND  (x1 = TRUE) AND  (x2 = TRUE) AND  (t0.Q = TRUE)) THEN 
        cstate58 := 6466; y0 := FALSE; y1 := FALSE; t0_start := TRUE; t0_up := FALSE; 
    ELSIF ((x0 = TRUE) AND  (x1 = FALSE) AND  (x2 = FALSE) AND  (t0.Q = FALSE)) THEN 
        cstate58 := 2120; y0 := FALSE; y1 := FALSE; t0_start := FALSE; 
    ELSIF ((x0 = TRUE) AND  (x1 = FALSE) AND  (x2 = FALSE) AND  (t0.Q = TRUE)) THEN 
        cstate58 := 2114; y0 := FALSE; y1 := FALSE; t0_start := FALSE; 
    ELSIF ((x0 = TRUE) AND  (x1 = FALSE) AND  (x2 = TRUE) AND  (t0.Q = FALSE)) THEN 
        cstate58 := 2760; y0 := FALSE; y1 := FALSE; t0_start := TRUE; t0_up := FALSE; 
    ELSIF ((x0 = TRUE) AND  (x1 = FALSE) AND  (x2 = TRUE) AND  (t0.Q = TRUE)) THEN 
        cstate58 := 2754; y0 := FALSE; y1 := FALSE; t0_start := TRUE; t0_up := FALSE; 
    ELSIF ((x0 = TRUE) AND  (x1 = TRUE) AND  (x2 = FALSE) AND  (t0.Q = FALSE)) THEN 
        cstate58 := 2630; y0 := FALSE; y1 := FALSE; t0_start := FALSE; 
    ELSIF ((x0 = TRUE) AND  (x1 = TRUE) AND  (x2 = FALSE) AND  (t0.Q = TRUE)) THEN 
        cstate58 := 2626; y0 := FALSE; y1 := FALSE; t0_start := FALSE; 
    ELSIF ((x0 = TRUE) AND  (x1 = TRUE) AND  (x2 = TRUE) AND  (t0.Q = FALSE)) THEN 
        cstate58 := 2566; y0 := FALSE; y1 := FALSE; t0_start := TRUE; t0_up := FALSE; 
    ELSIF ((x0 = TRUE) AND  (x1 = TRUE) AND  (x2 = TRUE) AND  (t0.Q = TRUE)) THEN 
        cstate58 := 2562; y0 := FALSE; y1 := FALSE; t0_start := TRUE; t0_up := FALSE; 
    END_IF;
2566:
    IF ((x0 = FALSE) AND  (x1 = FALSE) AND  (x2 = FALSE) AND  (t0.Q = FALSE)) THEN 
        cstate58 := 6404; y0 := FALSE; y1 := FALSE; t0_start := FALSE; 
    ELSIF ((x0 = FALSE) AND  (x1 = FALSE) AND  (x2 = FALSE) AND  (t0.Q = TRUE)) THEN 
        cstate58 := 6350; y0 := FALSE; y1 := TRUE; t0_start := FALSE; 
    ELSIF ((x0 = FALSE) AND  (x1 = FALSE) AND  (x2 = TRUE) AND  (t0.Q = FALSE)) THEN 
        cstate58 := 6468; y0 := FALSE; y1 := FALSE; t0_start := FALSE; 
    ELSIF ((x0 = FALSE) AND  (x1 = FALSE) AND  (x2 = TRUE) AND  (t0.Q = TRUE)) THEN 
        cstate58 := 6542; y0 := FALSE; y1 := TRUE; t0_start := FALSE; 
    ELSIF ((x0 = FALSE) AND  (x1 = TRUE) AND  (x2 = FALSE) AND  (t0.Q = FALSE)) THEN 
        cstate58 := 6404; y0 := FALSE; y1 := FALSE; t0_start := FALSE; 
    ELSIF ((x0 = FALSE) AND  (x1 = TRUE) AND  (x2 = FALSE) AND  (t0.Q = TRUE)) THEN 
        cstate58 := 6338; y0 := FALSE; y1 := FALSE; t0_start := FALSE; 
    ELSIF ((x0 = FALSE) AND  (x1 = TRUE) AND  (x2 = TRUE) AND  (t0.Q = FALSE)) THEN 
        cstate58 := 6468; y0 := FALSE; y1 := FALSE; t0_start := FALSE; 
    ELSIF ((x0 = FALSE) AND  (x1 = TRUE) AND  (x2 = TRUE) AND  (t0.Q = TRUE)) THEN 
        cstate58 := 6530; y0 := FALSE; y1 := FALSE; t0_start := FALSE; 
    ELSIF ((x0 = TRUE) AND  (x1 = FALSE) AND  (x2 = FALSE) AND  (t0.Q = FALSE)) THEN 
        cstate58 := 2184; y0 := FALSE; y1 := FALSE; t0_start := FALSE; 
    ELSIF ((x0 = TRUE) AND  (x1 = FALSE) AND  (x2 = FALSE) AND  (t0.Q = TRUE)) THEN 
        cstate58 := 2114; y0 := FALSE; y1 := FALSE; t0_start := FALSE; 
    ELSIF ((x0 = TRUE) AND  (x1 = FALSE) AND  (x2 = TRUE) AND  (t0.Q = FALSE)) THEN 
        cstate58 := 2760; y0 := FALSE; y1 := FALSE; t0_start := FALSE; 
    ELSIF ((x0 = TRUE) AND  (x1 = FALSE) AND  (x2 = TRUE) AND  (t0.Q = TRUE)) THEN 
        cstate58 := 2818; y0 := FALSE; y1 := FALSE; t0_start := FALSE; 
    ELSIF ((x0 = TRUE) AND  (x1 = TRUE) AND  (x2 = FALSE) AND  (t0.Q = FALSE)) THEN 
        cstate58 := 2694; y0 := FALSE; y1 := FALSE; t0_start := FALSE; 
    ELSIF ((x0 = TRUE) AND  (x1 = TRUE) AND  (x2 = FALSE) AND  (t0.Q = TRUE)) THEN 
        cstate58 := 2626; y0 := FALSE; y1 := FALSE; t0_start := FALSE; 
    ELSIF ((x0 = TRUE) AND  (x1 = TRUE) AND  (x2 = TRUE) AND  (t0.Q = FALSE)) THEN 
        cstate58 := 2566; y0 := FALSE; y1 := FALSE; t0_start := FALSE; 
    ELSIF ((x0 = TRUE) AND  (x1 = TRUE) AND  (x2 = TRUE) AND  (t0.Q = TRUE)) THEN 
        cstate58 := 2498; y0 := FALSE; y1 := FALSE; t0_start := FALSE; 
    END_IF;
4168:
    IF ((x0 = FALSE) AND  ( TRUE ) AND  (x2 = FALSE) AND  (t0.Q = FALSE)) THEN 
        cstate58 := 8388; y0 := TRUE; y1 := FALSE; t0_start := FALSE; 
    ELSIF ((x0 = FALSE) AND  ( TRUE ) AND  (x2 = FALSE) AND  (t0.Q = TRUE)) THEN 
        cstate58 := 8386; y0 := TRUE; y1 := FALSE; t0_start := FALSE; 
    ELSIF ((x0 = FALSE) AND  (x1 = FALSE) AND  (x2 = TRUE) AND  (t0.Q = FALSE)) THEN 
        cstate58 := 6468; y0 := FALSE; y1 := FALSE; t0_start := TRUE; t0_up := FALSE; 
    ELSIF ((x0 = FALSE) AND  (x1 = FALSE) AND  (x2 = TRUE) AND  (t0.Q = TRUE)) THEN 
        cstate58 := 6484; y0 := FALSE; y1 := TRUE; t0_start := TRUE; t0_up := FALSE; 
    ELSIF ((x0 = FALSE) AND  (x1 = TRUE) AND  (x2 = TRUE) AND  (t0.Q = FALSE)) THEN 
        cstate58 := 6468; y0 := FALSE; y1 := FALSE; t0_start := TRUE; t0_up := FALSE; 
    ELSIF ((x0 = FALSE) AND  (x1 = TRUE) AND  (x2 = TRUE) AND  (t0.Q = TRUE)) THEN 
        cstate58 := 6466; y0 := FALSE; y1 := FALSE; t0_start := TRUE; t0_up := FALSE; 
    ELSIF ((x0 = TRUE) AND  (x1 = FALSE) AND  (x2 = FALSE) AND  (t0.Q = FALSE)) THEN 
        cstate58 := 4168; y0 := TRUE; y1 := FALSE; t0_start := FALSE; 
    ELSIF ((x0 = TRUE) AND  (x1 = FALSE) AND  (x2 = FALSE) AND  (t0.Q = TRUE)) THEN 
        cstate58 := 4162; y0 := TRUE; y1 := FALSE; t0_start := FALSE; 
    ELSIF ((x0 = TRUE) AND  (x1 = FALSE) AND  (x2 = TRUE) AND  (t0.Q = FALSE)) THEN 
        cstate58 := 2760; y0 := FALSE; y1 := FALSE; t0_start := TRUE; t0_up := FALSE; 
    ELSIF ((x0 = TRUE) AND  (x1 = FALSE) AND  (x2 = TRUE) AND  (t0.Q = TRUE)) THEN 
        cstate58 := 2754; y0 := FALSE; y1 := FALSE; t0_start := TRUE; t0_up := FALSE; 
    ELSIF ((x0 = TRUE) AND  (x1 = TRUE) AND  (x2 = FALSE) AND  (t0.Q = FALSE)) THEN 
        cstate58 := 4678; y0 := TRUE; y1 := FALSE; t0_start := FALSE; 
    ELSIF ((x0 = TRUE) AND  (x1 = TRUE) AND  (x2 = FALSE) AND  (t0.Q = TRUE)) THEN 
        cstate58 := 4674; y0 := TRUE; y1 := FALSE; t0_start := FALSE; 
    ELSIF ((x0 = TRUE) AND  (x1 = TRUE) AND  (x2 = TRUE) AND  (t0.Q = FALSE)) THEN 
        cstate58 := 2566; y0 := FALSE; y1 := FALSE; t0_start := TRUE; t0_up := FALSE; 
    ELSIF ((x0 = TRUE) AND  (x1 = TRUE) AND  (x2 = TRUE) AND  (t0.Q = TRUE)) THEN 
        cstate58 := 2562; y0 := FALSE; y1 := FALSE; t0_start := TRUE; t0_up := FALSE; 
    END_IF;
2562:
    IF ((x0 = FALSE) AND  (x1 = FALSE) AND  (x2 = FALSE) AND  (t0.Q = FALSE)) THEN 
        cstate58 := 6404; y0 := FALSE; y1 := FALSE; t0_start := FALSE; 
    ELSIF ((x0 = FALSE) AND  (x1 = FALSE) AND  (x2 = FALSE) AND  (t0.Q = TRUE)) THEN 
        cstate58 := 6338; y0 := FALSE; y1 := FALSE; t0_start := FALSE; 
    ELSIF ((x0 = FALSE) AND  (x1 = FALSE) AND  (x2 = TRUE) AND  (t0.Q = FALSE)) THEN 
        cstate58 := 6468; y0 := FALSE; y1 := FALSE; t0_start := FALSE; 
    ELSIF ((x0 = FALSE) AND  (x1 = FALSE) AND  (x2 = TRUE) AND  (t0.Q = TRUE)) THEN 
        cstate58 := 6530; y0 := FALSE; y1 := FALSE; t0_start := FALSE; 
    ELSIF ((x0 = FALSE) AND  (x1 = TRUE) AND  (x2 = FALSE) AND  (t0.Q = FALSE)) THEN 
        cstate58 := 6404; y0 := FALSE; y1 := FALSE; t0_start := FALSE; 
    ELSIF ((x0 = FALSE) AND  (x1 = TRUE) AND  (x2 = FALSE) AND  (t0.Q = TRUE)) THEN 
        cstate58 := 6338; y0 := FALSE; y1 := FALSE; t0_start := FALSE; 
    ELSIF ((x0 = FALSE) AND  (x1 = TRUE) AND  (x2 = TRUE) AND  (t0.Q = FALSE)) THEN 
        cstate58 := 6468; y0 := FALSE; y1 := FALSE; t0_start := FALSE; 
    ELSIF ((x0 = FALSE) AND  (x1 = TRUE) AND  (x2 = TRUE) AND  (t0.Q = TRUE)) THEN 
        cstate58 := 6530; y0 := FALSE; y1 := FALSE; t0_start := FALSE; 
    ELSIF ((x0 = TRUE) AND  (x1 = FALSE) AND  (x2 = FALSE) AND  (t0.Q = FALSE)) THEN 
        cstate58 := 2184; y0 := FALSE; y1 := FALSE; t0_start := FALSE; 
    ELSIF ((x0 = TRUE) AND  (x1 = FALSE) AND  (x2 = FALSE) AND  (t0.Q = TRUE)) THEN 
        cstate58 := 2114; y0 := FALSE; y1 := FALSE; t0_start := FALSE; 
    ELSIF ((x0 = TRUE) AND  (x1 = FALSE) AND  (x2 = TRUE) AND  (t0.Q = FALSE)) THEN 
        cstate58 := 2760; y0 := FALSE; y1 := FALSE; t0_start := FALSE; 
    ELSIF ((x0 = TRUE) AND  (x1 = FALSE) AND  (x2 = TRUE) AND  (t0.Q = TRUE)) THEN 
        cstate58 := 2818; y0 := FALSE; y1 := FALSE; t0_start := FALSE; 
    ELSIF ((x0 = TRUE) AND  (x1 = TRUE) AND  (x2 = FALSE) AND  (t0.Q = FALSE)) THEN 
        cstate58 := 2694; y0 := FALSE; y1 := FALSE; t0_start := FALSE; 
    ELSIF ((x0 = TRUE) AND  (x1 = TRUE) AND  (x2 = FALSE) AND  (t0.Q = TRUE)) THEN 
        cstate58 := 2626; y0 := FALSE; y1 := FALSE; t0_start := FALSE; 
    ELSIF ((x0 = TRUE) AND  (x1 = TRUE) AND  (x2 = TRUE) AND  (t0.Q = FALSE)) THEN 
        cstate58 := 2566; y0 := FALSE; y1 := FALSE; t0_start := FALSE; 
    ELSIF ((x0 = TRUE) AND  (x1 = TRUE) AND  (x2 = TRUE) AND  (t0.Q = TRUE)) THEN 
        cstate58 := 2498; y0 := FALSE; y1 := FALSE; t0_start := FALSE; 
    END_IF;
7574:
    IF ((x0 = FALSE) AND  (x1 = FALSE) AND  (x2 = FALSE) AND  (t0.Q = FALSE)) THEN 
        cstate58 := 7382; y0 := FALSE; y1 := TRUE; t0_start := FALSE; 
    ELSIF ((x0 = FALSE) AND  (x1 = FALSE) AND  (x2 = FALSE) AND  (t0.Q = TRUE)) THEN 
        cstate58 := 7370; y0 := FALSE; y1 := TRUE; t0_start := FALSE; 
    ELSIF ((x0 = FALSE) AND  (x1 = FALSE) AND  (x2 = TRUE) AND  (t0.Q = FALSE)) THEN 
        cstate58 := 7574; y0 := FALSE; y1 := TRUE; t0_start := FALSE; 
    ELSIF ((x0 = FALSE) AND  (x1 = FALSE) AND  (x2 = TRUE) AND  (t0.Q = TRUE)) THEN 
        cstate58 := 7562; y0 := FALSE; y1 := TRUE; t0_start := FALSE; 
    ELSIF ((x0 = FALSE) AND  (x1 = TRUE) AND  (x2 = FALSE) AND  (t0.Q = FALSE)) THEN 
        cstate58 := 6340; y0 := FALSE; y1 := FALSE; t0_start := FALSE; 
    ELSIF ((x0 = FALSE) AND  (x1 = TRUE) AND  (x2 = FALSE) AND  (t0.Q = TRUE)) THEN 
        cstate58 := 6338; y0 := FALSE; y1 := FALSE; t0_start := FALSE; 
    ELSIF ((x0 = FALSE) AND  (x1 = TRUE) AND  (x2 = TRUE) AND  (t0.Q = FALSE)) THEN 
        cstate58 := 6532; y0 := FALSE; y1 := FALSE; t0_start := FALSE; 
    ELSIF ((x0 = FALSE) AND  (x1 = TRUE) AND  (x2 = TRUE) AND  (t0.Q = TRUE)) THEN 
        cstate58 := 6530; y0 := FALSE; y1 := FALSE; t0_start := FALSE; 
    ELSIF ((x0 = TRUE) AND  (x1 = FALSE) AND  (x2 = FALSE) AND  (t0.Q = FALSE)) THEN 
        cstate58 := 5192; y0 := TRUE; y1 := FALSE; t0_start := FALSE; 
    ELSIF ((x0 = TRUE) AND  (x1 = FALSE) AND  (x2 = FALSE) AND  (t0.Q = TRUE)) THEN 
        cstate58 := 5186; y0 := TRUE; y1 := FALSE; t0_start := FALSE; 
    ELSIF ((x0 = TRUE) AND  (x1 = FALSE) AND  (x2 = TRUE) AND  (t0.Q = FALSE)) THEN 
        cstate58 := 3848; y0 := FALSE; y1 := FALSE; t0_start := FALSE; 
    ELSIF ((x0 = TRUE) AND  (x1 = FALSE) AND  (x2 = TRUE) AND  (t0.Q = TRUE)) THEN 
        cstate58 := 3842; y0 := FALSE; y1 := FALSE; t0_start := FALSE; 
    ELSIF ((x0 = TRUE) AND  (x1 = TRUE) AND  (x2 = FALSE) AND  (t0.Q = FALSE)) THEN 
        cstate58 := 4678; y0 := TRUE; y1 := FALSE; t0_start := FALSE; 
    ELSIF ((x0 = TRUE) AND  (x1 = TRUE) AND  (x2 = FALSE) AND  (t0.Q = TRUE)) THEN 
        cstate58 := 4674; y0 := TRUE; y1 := FALSE; t0_start := FALSE; 
    ELSIF ((x0 = TRUE) AND  (x1 = TRUE) AND  (x2 = TRUE) AND  (t0.Q = FALSE)) THEN 
        cstate58 := 2502; y0 := FALSE; y1 := FALSE; t0_start := FALSE; 
    ELSIF ((x0 = TRUE) AND  (x1 = TRUE) AND  (x2 = TRUE) AND  (t0.Q = TRUE)) THEN 
        cstate58 := 2498; y0 := FALSE; y1 := FALSE; t0_start := FALSE; 
    END_IF;
5186:
    IF ((x0 = FALSE) AND  (x1 = FALSE) AND  (x2 = FALSE) AND  (t0.Q = FALSE)) THEN 
        cstate58 := 9412; y0 := TRUE; y1 := FALSE; t0_start := FALSE; 
    ELSIF ((x0 = FALSE) AND  (x1 = FALSE) AND  (x2 = FALSE) AND  (t0.Q = TRUE)) THEN 
        cstate58 := 9410; y0 := TRUE; y1 := FALSE; t0_start := FALSE; 
    ELSIF ((x0 = FALSE) AND  (x1 = FALSE) AND  (x2 = TRUE) AND  (t0.Q = FALSE)) THEN 
        cstate58 := 7492; y0 := FALSE; y1 := FALSE; t0_start := TRUE; t0_up := FALSE; 
    ELSIF ((x0 = FALSE) AND  (x1 = FALSE) AND  (x2 = TRUE) AND  (t0.Q = TRUE)) THEN 
        cstate58 := 7490; y0 := FALSE; y1 := FALSE; t0_start := TRUE; t0_up := FALSE; 
    ELSIF ((x0 = FALSE) AND  (x1 = TRUE) AND  (x2 = FALSE) AND  (t0.Q = FALSE)) THEN 
        cstate58 := 8388; y0 := TRUE; y1 := FALSE; t0_start := FALSE; 
    ELSIF ((x0 = FALSE) AND  (x1 = TRUE) AND  (x2 = FALSE) AND  (t0.Q = TRUE)) THEN 
        cstate58 := 8386; y0 := TRUE; y1 := FALSE; t0_start := FALSE; 
    ELSIF ((x0 = FALSE) AND  (x1 = TRUE) AND  (x2 = TRUE) AND  (t0.Q = FALSE)) THEN 
        cstate58 := 6468; y0 := FALSE; y1 := FALSE; t0_start := TRUE; t0_up := FALSE; 
    ELSIF ((x0 = FALSE) AND  (x1 = TRUE) AND  (x2 = TRUE) AND  (t0.Q = TRUE)) THEN 
        cstate58 := 6466; y0 := FALSE; y1 := FALSE; t0_start := TRUE; t0_up := FALSE; 
    ELSIF ((x0 = TRUE) AND  (x1 = FALSE) AND  (x2 = FALSE) AND  (t0.Q = FALSE)) THEN 
        cstate58 := 5192; y0 := TRUE; y1 := FALSE; t0_start := FALSE; 
    ELSIF ((x0 = TRUE) AND  (x1 = FALSE) AND  (x2 = FALSE) AND  (t0.Q = TRUE)) THEN 
        cstate58 := 5186; y0 := TRUE; y1 := FALSE; t0_start := FALSE; 
    ELSIF ((x0 = TRUE) AND  (x1 = FALSE) AND  (x2 = TRUE) AND  (t0.Q = FALSE)) THEN 
        cstate58 := 3784; y0 := FALSE; y1 := FALSE; t0_start := TRUE; t0_up := FALSE; 
    ELSIF ((x0 = TRUE) AND  (x1 = FALSE) AND  (x2 = TRUE) AND  (t0.Q = TRUE)) THEN 
        cstate58 := 3778; y0 := FALSE; y1 := FALSE; t0_start := TRUE; t0_up := FALSE; 
    ELSIF ((x0 = TRUE) AND  (x1 = TRUE) AND  (x2 = FALSE) AND  (t0.Q = FALSE)) THEN 
        cstate58 := 4678; y0 := TRUE; y1 := FALSE; t0_start := FALSE; 
    ELSIF ((x0 = TRUE) AND  (x1 = TRUE) AND  (x2 = FALSE) AND  (t0.Q = TRUE)) THEN 
        cstate58 := 4674; y0 := TRUE; y1 := FALSE; t0_start := FALSE; 
    ELSIF ((x0 = TRUE) AND  (x1 = TRUE) AND  (x2 = TRUE) AND  (t0.Q = FALSE)) THEN 
        cstate58 := 2566; y0 := FALSE; y1 := FALSE; t0_start := TRUE; t0_up := FALSE; 
    ELSIF ((x0 = TRUE) AND  (x1 = TRUE) AND  (x2 = TRUE) AND  (t0.Q = TRUE)) THEN 
        cstate58 := 2562; y0 := FALSE; y1 := FALSE; t0_start := TRUE; t0_up := FALSE; 
    END_IF;
2498:
    IF ((x0 = FALSE) AND  (x1 = FALSE) AND  (x2 = FALSE) AND  (t0.Q = FALSE)) THEN 
        cstate58 := 6340; y0 := FALSE; y1 := FALSE; t0_start := FALSE; 
    ELSIF ((x0 = FALSE) AND  (x1 = FALSE) AND  (x2 = FALSE) AND  (t0.Q = TRUE)) THEN 
        cstate58 := 6338; y0 := FALSE; y1 := FALSE; t0_start := FALSE; 
    ELSIF ((x0 = FALSE) AND  (x1 = FALSE) AND  (x2 = TRUE) AND  (t0.Q = FALSE)) THEN 
        cstate58 := 6532; y0 := FALSE; y1 := FALSE; t0_start := FALSE; 
    ELSIF ((x0 = FALSE) AND  (x1 = FALSE) AND  (x2 = TRUE) AND  (t0.Q = TRUE)) THEN 
        cstate58 := 6530; y0 := FALSE; y1 := FALSE; t0_start := FALSE; 
    ELSIF ((x0 = FALSE) AND  (x1 = TRUE) AND  (x2 = FALSE) AND  (t0.Q = FALSE)) THEN 
        cstate58 := 6340; y0 := FALSE; y1 := FALSE; t0_start := FALSE; 
    ELSIF ((x0 = FALSE) AND  (x1 = TRUE) AND  (x2 = FALSE) AND  (t0.Q = TRUE)) THEN 
        cstate58 := 6338; y0 := FALSE; y1 := FALSE; t0_start := FALSE; 
    ELSIF ((x0 = FALSE) AND  (x1 = TRUE) AND  (x2 = TRUE) AND  (t0.Q = FALSE)) THEN 
        cstate58 := 6532; y0 := FALSE; y1 := FALSE; t0_start := FALSE; 
    ELSIF ((x0 = FALSE) AND  (x1 = TRUE) AND  (x2 = TRUE) AND  (t0.Q = TRUE)) THEN 
        cstate58 := 6530; y0 := FALSE; y1 := FALSE; t0_start := FALSE; 
    ELSIF ((x0 = TRUE) AND  (x1 = FALSE) AND  (x2 = FALSE) AND  (t0.Q = FALSE)) THEN 
        cstate58 := 2120; y0 := FALSE; y1 := FALSE; t0_start := FALSE; 
    ELSIF ((x0 = TRUE) AND  (x1 = FALSE) AND  (x2 = FALSE) AND  (t0.Q = TRUE)) THEN 
        cstate58 := 2114; y0 := FALSE; y1 := FALSE; t0_start := FALSE; 
    ELSIF ((x0 = TRUE) AND  (x1 = FALSE) AND  (x2 = TRUE) AND  (t0.Q = FALSE)) THEN 
        cstate58 := 2824; y0 := FALSE; y1 := FALSE; t0_start := FALSE; 
    ELSIF ((x0 = TRUE) AND  (x1 = FALSE) AND  (x2 = TRUE) AND  (t0.Q = TRUE)) THEN 
        cstate58 := 2818; y0 := FALSE; y1 := FALSE; t0_start := FALSE; 
    ELSIF ((x0 = TRUE) AND  (x1 = TRUE) AND  (x2 = FALSE) AND  (t0.Q = FALSE)) THEN 
        cstate58 := 2630; y0 := FALSE; y1 := FALSE; t0_start := FALSE; 
    ELSIF ((x0 = TRUE) AND  (x1 = TRUE) AND  (x2 = FALSE) AND  (t0.Q = TRUE)) THEN 
        cstate58 := 2626; y0 := FALSE; y1 := FALSE; t0_start := FALSE; 
    ELSIF ((x0 = TRUE) AND  (x1 = TRUE) AND  (x2 = TRUE) AND  (t0.Q = FALSE)) THEN 
        cstate58 := 2502; y0 := FALSE; y1 := FALSE; t0_start := FALSE; 
    ELSIF ((x0 = TRUE) AND  (x1 = TRUE) AND  (x2 = TRUE) AND  (t0.Q = TRUE)) THEN 
        cstate58 := 2498; y0 := FALSE; y1 := FALSE; t0_start := FALSE; 
    END_IF;
6340:
    IF ((x0 = FALSE) AND  (x1 = FALSE) AND  (x2 = FALSE) AND  (t0.Q = FALSE)) THEN 
        cstate58 := 6340; y0 := FALSE; y1 := FALSE; t0_start := FALSE; 
    ELSIF ((x0 = FALSE) AND  (x1 = FALSE) AND  (x2 = FALSE) AND  (t0.Q = TRUE)) THEN 
        cstate58 := 6346; y0 := FALSE; y1 := TRUE; t0_start := FALSE; 
    ELSIF ((x0 = FALSE) AND  (x1 = FALSE) AND  (x2 = TRUE) AND  (t0.Q = FALSE)) THEN 
        cstate58 := 6468; y0 := FALSE; y1 := FALSE; t0_start := TRUE; t0_up := FALSE; 
    ELSIF ((x0 = FALSE) AND  (x1 = FALSE) AND  (x2 = TRUE) AND  (t0.Q = TRUE)) THEN 
        cstate58 := 6476; y0 := FALSE; y1 := TRUE; t0_start := TRUE; t0_up := FALSE; 
    ELSIF ((x0 = FALSE) AND  (x1 = TRUE) AND  (x2 = FALSE) AND  (t0.Q = FALSE)) THEN 
        cstate58 := 6340; y0 := FALSE; y1 := FALSE; t0_start := FALSE; 
    ELSIF ((x0 = FALSE) AND  (x1 = TRUE) AND  (x2 = FALSE) AND  (t0.Q = TRUE)) THEN 
        cstate58 := 6338; y0 := FALSE; y1 := FALSE; t0_start := FALSE; 
    ELSIF ((x0 = FALSE) AND  (x1 = TRUE) AND  (x2 = TRUE) AND  (t0.Q = FALSE)) THEN 
        cstate58 := 6468; y0 := FALSE; y1 := FALSE; t0_start := TRUE; t0_up := FALSE; 
    ELSIF ((x0 = FALSE) AND  (x1 = TRUE) AND  (x2 = TRUE) AND  (t0.Q = TRUE)) THEN 
        cstate58 := 6466; y0 := FALSE; y1 := FALSE; t0_start := TRUE; t0_up := FALSE; 
    ELSIF ((x0 = TRUE) AND  (x1 = FALSE) AND  (x2 = FALSE) AND  (t0.Q = FALSE)) THEN 
        cstate58 := 4168; y0 := TRUE; y1 := FALSE; t0_start := FALSE; 
    ELSIF ((x0 = TRUE) AND  (x1 = FALSE) AND  (x2 = FALSE) AND  (t0.Q = TRUE)) THEN 
        cstate58 := 4162; y0 := TRUE; y1 := FALSE; t0_start := FALSE; 
    ELSIF ((x0 = TRUE) AND  (x1 = FALSE) AND  (x2 = TRUE) AND  (t0.Q = FALSE)) THEN 
        cstate58 := 2760; y0 := FALSE; y1 := FALSE; t0_start := TRUE; t0_up := FALSE; 
    ELSIF ((x0 = TRUE) AND  (x1 = FALSE) AND  (x2 = TRUE) AND  (t0.Q = TRUE)) THEN 
        cstate58 := 2754; y0 := FALSE; y1 := FALSE; t0_start := TRUE; t0_up := FALSE; 
    ELSIF ((x0 = TRUE) AND  (x1 = TRUE) AND  (x2 = FALSE) AND  (t0.Q = FALSE)) THEN 
        cstate58 := 4678; y0 := TRUE; y1 := FALSE; t0_start := FALSE; 
    ELSIF ((x0 = TRUE) AND  (x1 = TRUE) AND  (x2 = FALSE) AND  (t0.Q = TRUE)) THEN 
        cstate58 := 4674; y0 := TRUE; y1 := FALSE; t0_start := FALSE; 
    ELSIF ((x0 = TRUE) AND  (x1 = TRUE) AND  (x2 = TRUE) AND  (t0.Q = FALSE)) THEN 
        cstate58 := 2566; y0 := FALSE; y1 := FALSE; t0_start := TRUE; t0_up := FALSE; 
    ELSIF ((x0 = TRUE) AND  (x1 = TRUE) AND  (x2 = TRUE) AND  (t0.Q = TRUE)) THEN 
        cstate58 := 2562; y0 := FALSE; y1 := FALSE; t0_start := TRUE; t0_up := FALSE; 
    END_IF;
6346:
    IF ((x0 = FALSE) AND  (x1 = FALSE) AND  (x2 = FALSE) AND  (t0.Q = FALSE)) THEN 
        cstate58 := 6358; y0 := FALSE; y1 := TRUE; t0_start := FALSE; 
    ELSIF ((x0 = FALSE) AND  (x1 = FALSE) AND  (x2 = FALSE) AND  (t0.Q = TRUE)) THEN 
        cstate58 := 6346; y0 := FALSE; y1 := TRUE; t0_start := FALSE; 
    ELSIF ((x0 = FALSE) AND  (x1 = FALSE) AND  (x2 = TRUE) AND  (t0.Q = FALSE)) THEN 
        cstate58 := 6488; y0 := FALSE; y1 := TRUE; t0_start := TRUE; t0_up := FALSE; 
    ELSIF ((x0 = FALSE) AND  (x1 = FALSE) AND  (x2 = TRUE) AND  (t0.Q = TRUE)) THEN 
        cstate58 := 6476; y0 := FALSE; y1 := TRUE; t0_start := TRUE; t0_up := FALSE; 
    ELSIF ((x0 = FALSE) AND  (x1 = TRUE) AND  (x2 = FALSE) AND  (t0.Q = FALSE)) THEN 
        cstate58 := 6340; y0 := FALSE; y1 := FALSE; t0_start := FALSE; 
    ELSIF ((x0 = FALSE) AND  (x1 = TRUE) AND  (x2 = FALSE) AND  (t0.Q = TRUE)) THEN 
        cstate58 := 6338; y0 := FALSE; y1 := FALSE; t0_start := FALSE; 
    ELSIF ((x0 = FALSE) AND  (x1 = TRUE) AND  (x2 = TRUE) AND  (t0.Q = FALSE)) THEN 
        cstate58 := 6468; y0 := FALSE; y1 := FALSE; t0_start := TRUE; t0_up := FALSE; 
    ELSIF ((x0 = FALSE) AND  (x1 = TRUE) AND  (x2 = TRUE) AND  (t0.Q = TRUE)) THEN 
        cstate58 := 6466; y0 := FALSE; y1 := FALSE; t0_start := TRUE; t0_up := FALSE; 
    ELSIF ((x0 = TRUE) AND  (x1 = FALSE) AND  (x2 = FALSE) AND  (t0.Q = FALSE)) THEN 
        cstate58 := 4168; y0 := TRUE; y1 := FALSE; t0_start := FALSE; 
    ELSIF ((x0 = TRUE) AND  (x1 = FALSE) AND  (x2 = FALSE) AND  (t0.Q = TRUE)) THEN 
        cstate58 := 4162; y0 := TRUE; y1 := FALSE; t0_start := FALSE; 
    ELSIF ((x0 = TRUE) AND  (x1 = FALSE) AND  (x2 = TRUE) AND  (t0.Q = FALSE)) THEN 
        cstate58 := 2760; y0 := FALSE; y1 := FALSE; t0_start := TRUE; t0_up := FALSE; 
    ELSIF ((x0 = TRUE) AND  (x1 = FALSE) AND  (x2 = TRUE) AND  (t0.Q = TRUE)) THEN 
        cstate58 := 2754; y0 := FALSE; y1 := FALSE; t0_start := TRUE; t0_up := FALSE; 
    ELSIF ((x0 = TRUE) AND  (x1 = TRUE) AND  (x2 = FALSE) AND  (t0.Q = FALSE)) THEN 
        cstate58 := 4678; y0 := TRUE; y1 := FALSE; t0_start := FALSE; 
    ELSIF ((x0 = TRUE) AND  (x1 = TRUE) AND  (x2 = FALSE) AND  (t0.Q = TRUE)) THEN 
        cstate58 := 4674; y0 := TRUE; y1 := FALSE; t0_start := FALSE; 
    ELSIF ((x0 = TRUE) AND  (x1 = TRUE) AND  (x2 = TRUE) AND  (t0.Q = FALSE)) THEN 
        cstate58 := 2566; y0 := FALSE; y1 := FALSE; t0_start := TRUE; t0_up := FALSE; 
    ELSIF ((x0 = TRUE) AND  (x1 = TRUE) AND  (x2 = TRUE) AND  (t0.Q = TRUE)) THEN 
        cstate58 := 2562; y0 := FALSE; y1 := FALSE; t0_start := TRUE; t0_up := FALSE; 
    END_IF;
6538:
    IF ((x0 = FALSE) AND  (x1 = FALSE) AND  (x2 = FALSE) AND  (t0.Q = FALSE)) THEN 
        cstate58 := 6358; y0 := FALSE; y1 := TRUE; t0_start := FALSE; 
    ELSIF ((x0 = FALSE) AND  (x1 = FALSE) AND  (x2 = FALSE) AND  (t0.Q = TRUE)) THEN 
        cstate58 := 6346; y0 := FALSE; y1 := TRUE; t0_start := FALSE; 
    ELSIF ((x0 = FALSE) AND  (x1 = FALSE) AND  (x2 = TRUE) AND  (t0.Q = FALSE)) THEN 
        cstate58 := 6550; y0 := FALSE; y1 := TRUE; t0_start := FALSE; 
    ELSIF ((x0 = FALSE) AND  (x1 = FALSE) AND  (x2 = TRUE) AND  (t0.Q = TRUE)) THEN 
        cstate58 := 6538; y0 := FALSE; y1 := TRUE; t0_start := FALSE; 
    ELSIF ((x0 = FALSE) AND  (x1 = TRUE) AND  (x2 = FALSE) AND  (t0.Q = FALSE)) THEN 
        cstate58 := 6340; y0 := FALSE; y1 := FALSE; t0_start := FALSE; 
    ELSIF ((x0 = FALSE) AND  (x1 = TRUE) AND  (x2 = FALSE) AND  (t0.Q = TRUE)) THEN 
        cstate58 := 6338; y0 := FALSE; y1 := FALSE; t0_start := FALSE; 
    ELSIF ((x0 = FALSE) AND  (x1 = TRUE) AND  (x2 = TRUE) AND  (t0.Q = FALSE)) THEN 
        cstate58 := 6532; y0 := FALSE; y1 := FALSE; t0_start := FALSE; 
    ELSIF ((x0 = FALSE) AND  (x1 = TRUE) AND  (x2 = TRUE) AND  (t0.Q = TRUE)) THEN 
        cstate58 := 6530; y0 := FALSE; y1 := FALSE; t0_start := FALSE; 
    ELSIF ((x0 = TRUE) AND  (x1 = FALSE) AND  (x2 = FALSE) AND  (t0.Q = FALSE)) THEN 
        cstate58 := 4168; y0 := TRUE; y1 := FALSE; t0_start := FALSE; 
    ELSIF ((x0 = TRUE) AND  (x1 = FALSE) AND  (x2 = FALSE) AND  (t0.Q = TRUE)) THEN 
        cstate58 := 4162; y0 := TRUE; y1 := FALSE; t0_start := FALSE; 
    ELSIF ((x0 = TRUE) AND  (x1 = FALSE) AND  (x2 = TRUE) AND  (t0.Q = FALSE)) THEN 
        cstate58 := 2824; y0 := FALSE; y1 := FALSE; t0_start := FALSE; 
    ELSIF ((x0 = TRUE) AND  (x1 = FALSE) AND  (x2 = TRUE) AND  (t0.Q = TRUE)) THEN 
        cstate58 := 2818; y0 := FALSE; y1 := FALSE; t0_start := FALSE; 
    ELSIF ((x0 = TRUE) AND  (x1 = TRUE) AND  (x2 = FALSE) AND  (t0.Q = FALSE)) THEN 
        cstate58 := 4678; y0 := TRUE; y1 := FALSE; t0_start := FALSE; 
    ELSIF ((x0 = TRUE) AND  (x1 = TRUE) AND  (x2 = FALSE) AND  (t0.Q = TRUE)) THEN 
        cstate58 := 4674; y0 := TRUE; y1 := FALSE; t0_start := FALSE; 
    ELSIF ((x0 = TRUE) AND  (x1 = TRUE) AND  (x2 = TRUE) AND  (t0.Q = FALSE)) THEN 
        cstate58 := 2502; y0 := FALSE; y1 := FALSE; t0_start := FALSE; 
    ELSIF ((x0 = TRUE) AND  (x1 = TRUE) AND  (x2 = TRUE) AND  (t0.Q = TRUE)) THEN 
        cstate58 := 2498; y0 := FALSE; y1 := FALSE; t0_start := FALSE; 
    END_IF;
7570:
